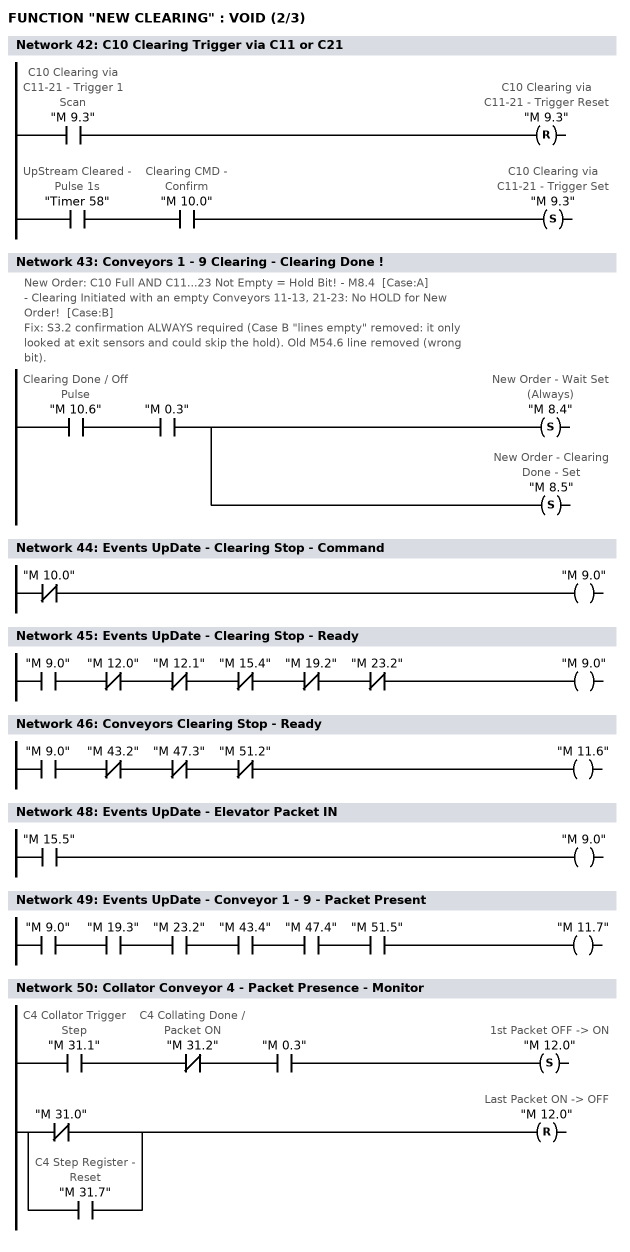

      A     "M 9.3"; // C10 Clearing via C11-21 - Trigger 1 Scan
      R     "M 9.3"; // C10 Clearing via C11-21 - Trigger Reset
//;
      A     "Timer 58"; // UpStream Cleared - Pulse 1s
      A     "M 10.0"; // Clearing CMD - Confirm
      S     "M 9.3"; // C10 Clearing via C11-21 - Trigger Set
NETWORK
TITLE =Conveyors 1 - 9 Clearing - Clearing Done !
//New Order: C10 Full AND C11...23 Not Empty = Hold Bit! - M8.4  [Case:A]
//
//- Clearing Initiated with an empty Conveyors 11-13, 21-23: No HOLD for New
//Order!  [Case:B]
//
//Fix: S3.2 confirmation ALWAYS required (Case B "lines empty" removed: it only
//looked at exit sensors and could skip the hold). Old M54.6 line removed (wrong
//bit).
      A     "M 10.6"; // Clearing Done / Off Pulse
      A     "M 0.3";
      S     "M 8.4"; // New Order - Wait Set (Always)
      S     "M 8.5"; // New Order - Clearing Done - Set
NETWORK
TITLE =Events UpDate - Clearing Stop - Command

      AN    "M 10.0";
      =     "M 9.0";
NETWORK
TITLE =Events UpDate - Clearing Stop - Ready

      A     "M 9.0";
      AN    "M 12.0";
      AN    "M 12.1";
      AN    "M 15.4";
      AN    "M 19.2";
      AN    "M 23.2";
      =     "M 9.0";
NETWORK
TITLE =Conveyors Clearing Stop - Ready

      A     "M 9.0";
      AN    "M 43.2";
      AN    "M 47.3";
      AN    "M 51.2";
      =     "M 11.6";
NETWORK
TITLE =New Order
//New Order : Start Filling Conveyors


NETWORK
TITLE =Events UpDate - Elevator Packet IN

      A     "M 15.5";
      =     "M 9.0";
NETWORK
TITLE =Events UpDate - Conveyor 1 - 9 - Packet Present

      A     "M 9.0";
      A     "M 19.3";
      A     "M 23.2";
      A     "M 43.4";
      A     "M 47.4";
      A     "M 51.5";
      =     "M 11.7";
NETWORK
TITLE =Collator Conveyor 4 - Packet Presence - Monitor

      A     "M 31.1"; // C4 Collator Trigger Step
      AN    "M 31.2"; // C4 Collating Done / Packet ON
      A     "M 0.3";
      S     "M 12.0"; // 1st Packet OFF -> ON
//;
      A(    ;
      ON    "M 31.0";
      O     "M 31.7"; // C4 Step Register - Reset
      )     ;
      R     "M 12.0"; // Last Packet ON -> OFF
NETWORK
TITLE =Collator Conveyor 10 - Packet Presence - Monitor
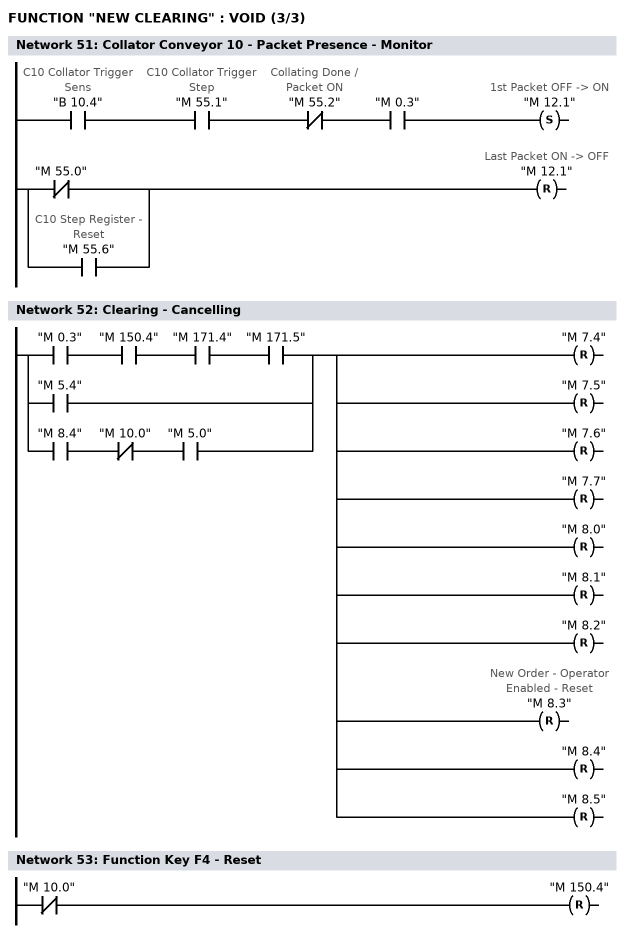

      A     "B 10.4"; // C10 Collator Trigger Sens
      A     "M 55.1"; // C10 Collator Trigger Step
      AN    "M 55.2"; // Collating Done / Packet ON
      A     "M 0.3";
      S     "M 12.1"; // 1st Packet OFF -> ON
//;
      A(    ;
      ON    "M 55.0";
      O     "M 55.6"; // C10 Step Register - Reset
      )     ;
      R     "M 12.1"; // Last Packet ON -> OFF
NETWORK
TITLE =Clearing - Cancelling

      A     "M 0.3";
      A     "M 150.4";
      A     "M 171.4";
      A     "M 171.5";
      O     "M 5.4";
      O(    ;
      A     "M 8.4";
      AN    "M 10.0";
      A     "M 5.0";
      )     ;
      R     "M 7.4";
      R     "M 7.5";
      R     "M 7.6";
      R     "M 7.7";
      R     "M 8.0";
      R     "M 8.1";
      R     "M 8.2";
      R     "M 8.3"; // New Order - Operator Enabled - Reset
      R     "M 8.4";
      R     "M 8.5";
NETWORK
TITLE =Function Key F4 - Reset

      AN    "M 10.0";
      R     "M 150.4";
END_FUNCTION

FUNCTION "NEW C0 + PUSHER 0" : VOID
TITLE =NEW FC912 (was FC1012) - Conveyor 0 & Pusher 0
NAME : 'Pos.1'
VERSION : 0.1


VAR_TEMP
  TIMER_RESET : BOOL ;
  MAIN_SERVICE_1_SW : BOOL ;
  CONV_0_SERVICE_FWD : BOOL ;
  CONV_0_SERVICE_REV : BOOL ;
  RESET_1 : BOOL ;
  RESET_2 : BOOL ;
  PUSHER_PUSH : BOOL ;
END_VAR
BEGIN
NETWORK
TITLE =Conveyor 0 - Service

      A     "HMI_DB".ALL_SERVICE_ENABLE_SW;
      A     "HMI_DB".CONVEYOR_0_SERVICE_SW;
      A     "HMI_DB".SERVICE_SW_1_STATUS;
      =     #MAIN_SERVICE_1_SW;
//;
      A     #MAIN_SERVICE_1_SW;
      O     "M 14.0";
      JNB   PUS0;
      A     "HMI_DB".HMI_ROLLER_TEST_FWD_SSW;
      FP    "FP 168.3";
      R     "HMI_DB".HMI_ROLLER_TEST_REV_SSW;
      =     #RESET_1;
//;
      A     "HMI_DB".HMI_ROLLER_TEST_REV_SSW;
      FP    "FP 168.4";
      R     "HMI_DB".HMI_ROLLER_TEST_FWD_SSW;
      =     #RESET_2;
//;
      A(    ;
      O     #RESET_1;
      O     #RESET_2;
      )     ;
      L     S5T#1S;
      SF    "Timer 110";
//;
      A     "HMI_DB".HMI_ROLLER_TEST_FWD_SSW;
      AN    "Timer 110";
      =     #CONV_0_SERVICE_FWD;
//;
      A     "HMI_DB".HMI_ROLLER_TEST_REV_SSW;
      AN    "Timer 110";
      =     #CONV_0_SERVICE_REV;
//;
      A     "HMI_DB".HMI_PUSHER_0_TEST_SSW;
      =     #PUSHER_PUSH;
//;
      AN    #MAIN_SERVICE_1_SW;
      R     "HMI_DB".HMI_ROLLER_TEST_FWD_SSW;
      R     "HMI_DB".HMI_ROLLER_TEST_REV_SSW;

PUS0: R     #CONV_0_SERVICE_FWD;
      R     #CONV_0_SERVICE_REV;
      R     #RESET_1;
      R     #RESET_2;
      R     #PUSHER_PUSH;
      FP    "FP 158.0";
      =     "M 14.0";
NETWORK
TITLE =Function Keys <F5 > on HMI - Reset
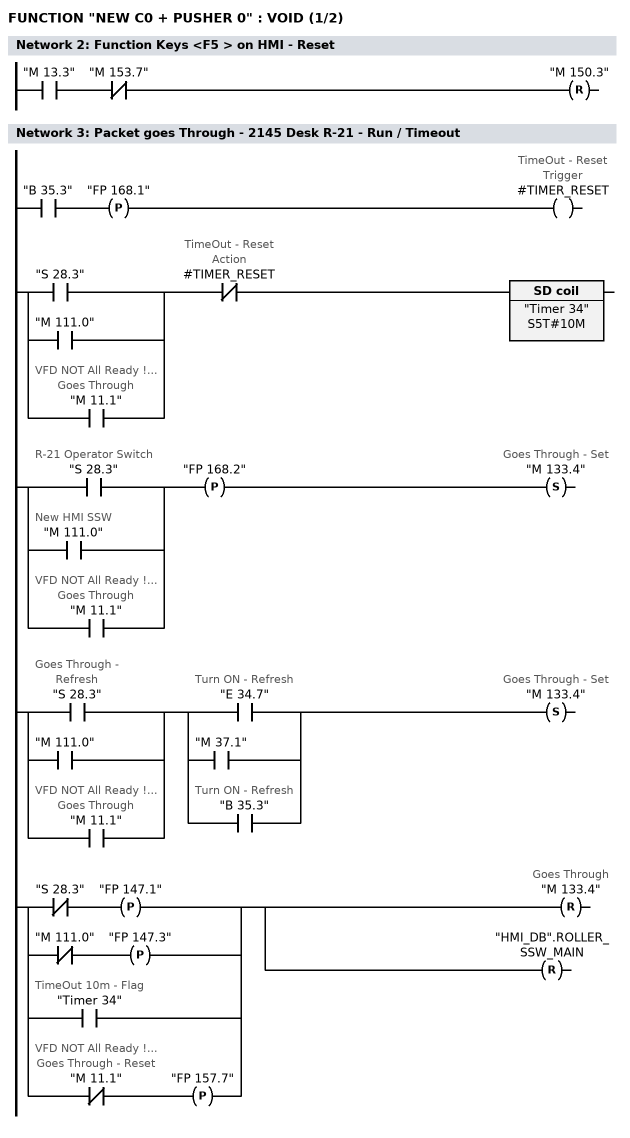

      A     "M 13.3";
      AN    "M 153.7";
      R     "M 150.3";
NETWORK
TITLE =Packet goes Through - 2145 Desk R-21 - Run / Timeout

      A     "B 35.3";
      FP    "FP 168.1";
      =     #TIMER_RESET; // TimeOut - Reset Trigger
//;
      A     "S 28.3";
      O     "M 111.0";
      O     "M 11.1"; // VFD NOT All Ready !... Goes Through
      AN    #TIMER_RESET; // TimeOut - Reset Action
      L     S5T#10M;
      SD    "Timer 34"; // TimeOut 10m
//;
      A     "S 28.3"; // R-21 Operator Switch
      O     "M 111.0"; // New HMI SSW
      O     "M 11.1"; // VFD NOT All Ready !... Goes Through
      FP    "FP 168.2"; // Turn ON - Pulse
      S     "M 133.4"; // Goes Through - Set
//;
      A     "S 28.3"; // Goes Through - Refresh
      O     "M 111.0";
      O     "M 11.1"; // VFD NOT All Ready !... Goes Through
      A(    ;
      O     "E 34.7"; // Turn ON - Refresh
      O     "M 37.1";
      O     "B 35.3"; // Turn ON - Refresh
      )     ;
      S     "M 133.4"; // Goes Through - Set
//;
      A(    ;
      O(    ;
      AN    "S 28.3";
      FP    "FP 147.1"; // Turn OFF - Pulse
      )     ;
      O(    ;
      AN    "M 111.0";
      FP    "FP 147.3"; // Turn OFF - Pulse
      O     "Timer 34"; // TimeOut 10m - Flag
      )     ;
      O(    ;
      AN    "M 11.1"; // VFD NOT All Ready !... Goes Through - Reset
      FP    "FP 157.7";
      )     ;
      )     ;
      R     "M 133.4"; // Goes Through
      R     "HMI_DB".ROLLER_SSW_MAIN;
NETWORK
TITLE =
//
//      A     "E 2.4"
//      S     "M 33.0"                    // Solid Detected ?
////;
//      A     "M 33.0"                    // Delay Timer - Start
//      L     S5T#300MS
//      SD    "Timer 26"                  // Debouncer 300mS
////;
//      A     "Timer 26"                  // Delayed Test Pulse
//      AN    "E 2.4"                     // Foul Detection
//      R     "M 33.0"                    // Not Detected !
////;
//      A     "Timer 26"                  // Delayed Test Pulse
//      A     "M 33.0"                    // Detection Comfirm !
//      =     "M 33.1"                    // Packet Height OK
//      R     "M 33.0"                    // Reset
//


NETWORK
TITLE =Packet Height - Sensing / Debouncing
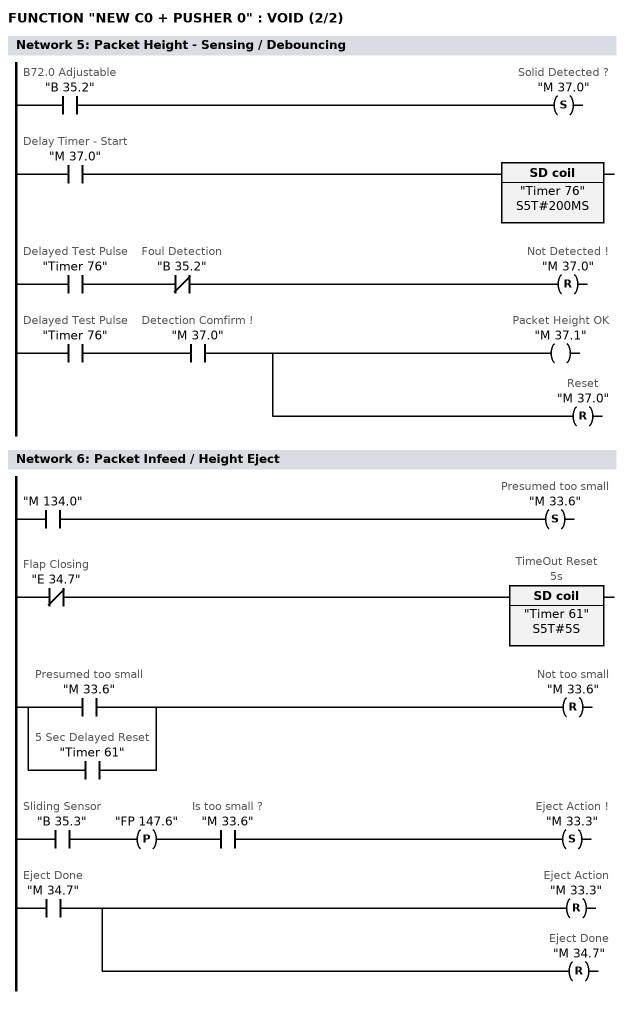

      A     "B 35.2"; // B72.0 Adjustable
      S     "M 37.0"; // Solid Detected ?
//;
      A     "M 37.0"; // Delay Timer - Start
      L     S5T#200MS;
      SD    "Timer 76"; // Debouncer 300mS
//;
      A     "Timer 76"; // Delayed Test Pulse
      AN    "B 35.2"; // Foul Detection
      R     "M 37.0"; // Not Detected !
//;
      A     "Timer 76"; // Delayed Test Pulse
      A     "M 37.0"; // Detection Comfirm !
      =     "M 37.1"; // Packet Height OK
      R     "M 37.0"; // Reset
NETWORK
TITLE =Packet Infeed / Height Eject

      A     "M 134.0";
      S     "M 33.6"; // Presumed too small
//;
      AN    "E 34.7"; // Flap Closing
      L     S5T#5S; // TimeOut Reset 5s
      SD    "Timer 61";
//;
      A     "M 33.6"; // Presumed too small
//    A     "M 33.1"                    // Packet Height OK ?
      O     "Timer 61"; // 5 Sec Delayed Reset
      R     "M 33.6"; // Not too small
//;
      A     "B 35.3"; // Sliding Sensor
      FP    "FP 147.6";
      A     "M 33.6"; // Is too small ?
      S     "M 33.3"; // Eject Action !
//;
      A     "M 34.7"; // Eject Done
      R     "M 33.3"; // Eject Action
      R     "M 34.7"; // Eject Done
NETWORK
TITLE =Eject Comfirmation

      A     "M 13.0";
      JNB   OUT1;

      A     "B 35.3";
      AN    "M 132.6"; // Not Triggered by Pusher
      S     "M 34.3"; // Eject Step 1
//;
      A     "B 35.4";
      AN    "M 132.6"; // Not Triggered by Pusher
      S     "M 34.4"; // Eject Step 2
//;
      A     "K 62.0"; // Conveyor 0 - Running
      A     "M 153.7";
      A     "M 34.3"; // Eject Step 1
      A     "M 34.4"; // Eject Step 2
      S     "M 34.5"; // Eject Step 3
//;
      A     "M 34.5"; // Eject Step 3
      AN    "B 35.4"; // Eject Step 4
      S     "M 34.7"; // Eject Done
      R     "M 34.3"; // Eject Step 1 - Reset
      R     "M 34.4"; // Eject Step 2 - Reset
      R     "M 34.5"; // Eject Step 3 - Reset
      R     "M 33.3"; // Eject Action - Reset
//;
      A     "M 132.5"; // Reset with Pusher Extend
      A     "B 35.4";
      R     "M 34.3"; // Eject Step 1 - Reset
      R     "M 34.4"; // Eject Step 2 - Reset
      R     "M 34.5"; // Eject Step 3 - Reset
      R     "M 33.3"; // Eject Action - Reset

OUT1: CLR   ;
NETWORK
TITLE =Packet goes Through - Conveyor 0 Man Run - LAUER F5
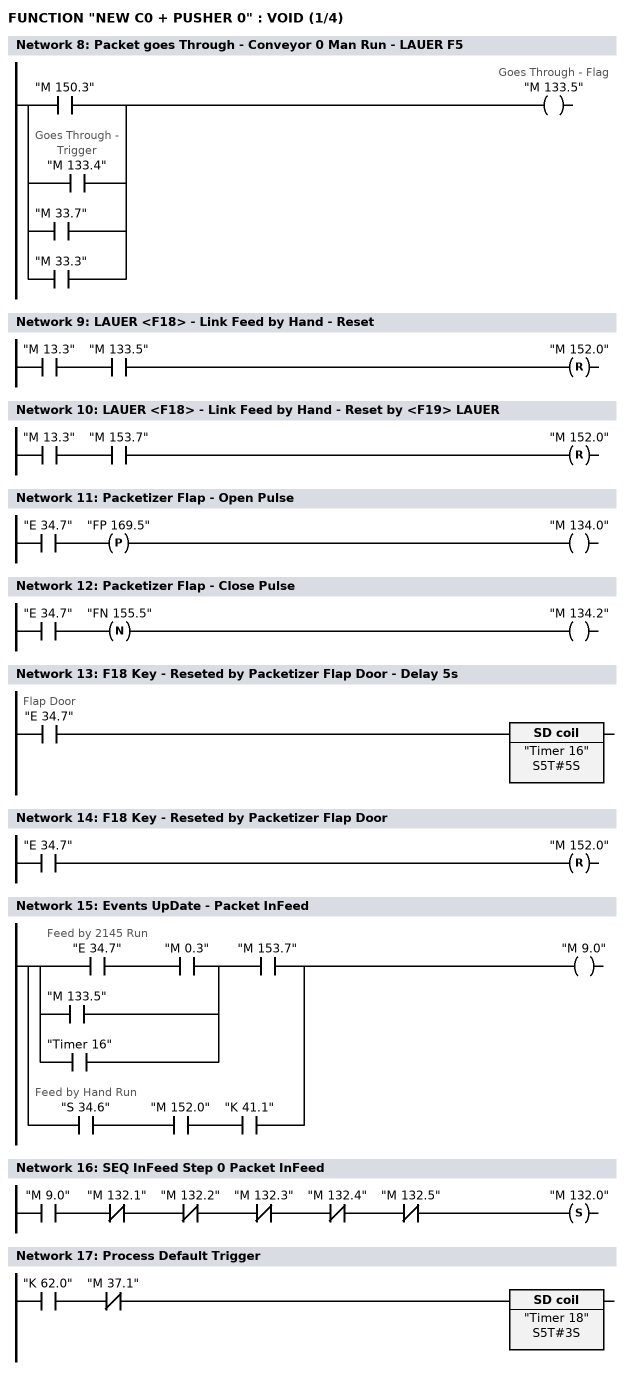

      O     "M 150.3";
      O     "M 133.4"; // Goes Through - Trigger
      O     "M 33.7";
      O     "M 33.3";
      =     "M 133.5"; // Goes Through - Flag
NETWORK
TITLE =LAUER <F18> - Link Feed by Hand - Reset

      A     "M 13.3";
      A     "M 133.5";
      R     "M 152.0";
NETWORK
TITLE =LAUER <F18> - Link Feed by Hand - Reset by <F19> LAUER

      A     "M 13.3";
      A     "M 153.7";
      R     "M 152.0";
NETWORK
TITLE =Packetizer Flap - Open Pulse

      A     "E 34.7";
      FP    "FP 169.5";
      =     "M 134.0";
NETWORK
TITLE =Packetizer Flap - Close Pulse

      A     "E 34.7";
      FN    "FN 155.5";
      =     "M 134.2";
NETWORK
TITLE =F18 Key - Reseted by Packetizer Flap Door - Delay 5s

      A     "E 34.7"; // Flap Door
      L     S5T#5S;
      SD    "Timer 16"; // Setup Mode Trigger
NETWORK
TITLE =F18 Key - Reseted by Packetizer Flap Door

      A     "E 34.7";
      R     "M 152.0";
NETWORK
TITLE =Events UpDate - Packet InFeed

      A(    ;
      A     "E 34.7"; // Feed by 2145 Run
      A     "M 0.3";
      O     "M 133.5";
      O     "Timer 16";
      A     "M 153.7";
      O     ;
      A     "S 34.6"; // Feed by Hand Run
      A     "M 152.0";
      A     "K 41.1";
      )     ;
      =     "M 9.0";
NETWORK
TITLE =SEQ InFeed Step 0 Packet InFeed

      A     "M 9.0";
      AN    "M 132.1";
      AN    "M 132.2";
      AN    "M 132.3";
      AN    "M 132.4";
      AN    "M 132.5";
      S     "M 132.0";
NETWORK
TITLE =Process Default Trigger

      A     "K 62.0";
      AN    "M 37.1";
      L     S5T#3S;
      SD    "Timer 18";
NETWORK
TITLE =Events UpDate
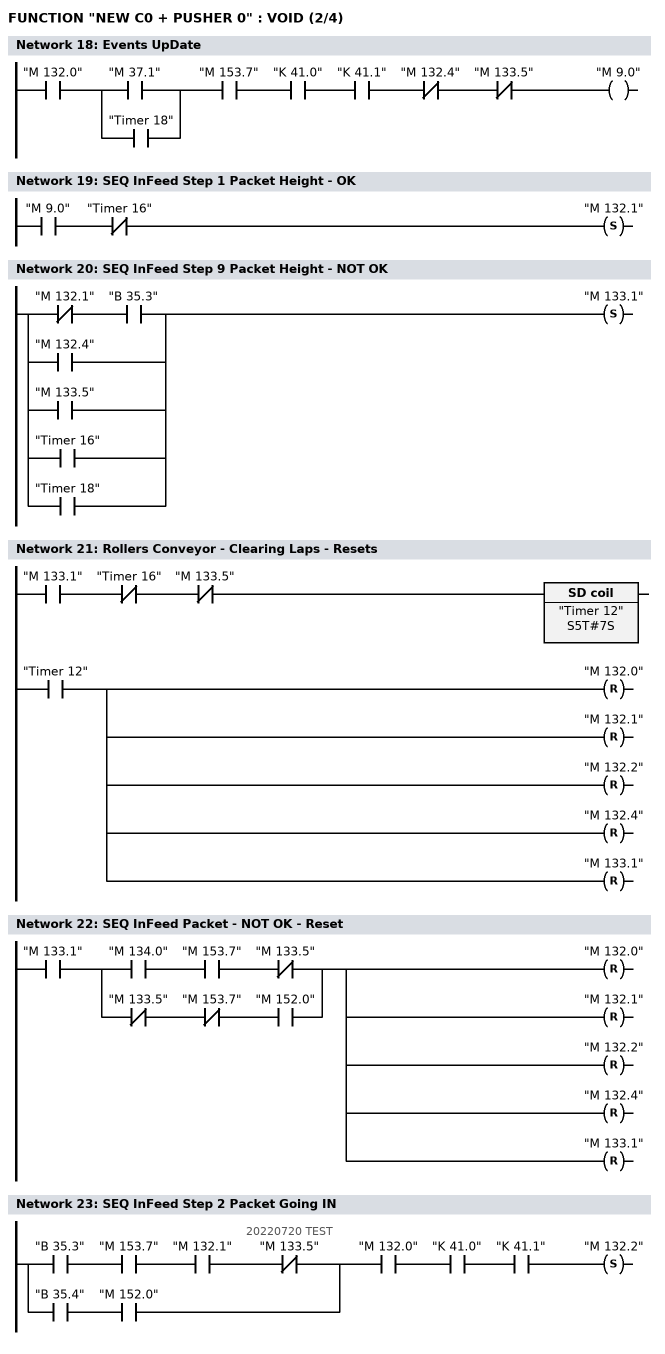

      A     "M 132.0";
      A(    ;
      O     "M 37.1";
      O     "Timer 18";
      )     ;
      A     "M 153.7";
      A     "K 41.0";
      A     "K 41.1";
      AN    "M 132.4";
      AN    "M 133.5";
      =     "M 9.0";
NETWORK
TITLE =SEQ InFeed Step 1 Packet Height - OK

      A     "M 9.0";
      AN    "Timer 16";
      S     "M 132.1";
NETWORK
TITLE =SEQ InFeed Step 9 Packet Height - NOT OK

      AN    "M 132.1";
      A     "B 35.3";
      O     "M 132.4";
      O     "M 133.5";
      O     "Timer 16";
      O     "Timer 18";
      S     "M 133.1";
NETWORK
TITLE =Rollers Conveyor - Clearing Laps - Resets

      A     "M 133.1";
      AN    "Timer 16";
      AN    "M 133.5";
      L     S5T#7S;
      SD    "Timer 12";
//;
      A     "Timer 12";
      R     "M 132.0";
      R     "M 132.1";
      R     "M 132.2";
      R     "M 132.4";
      R     "M 133.1";
NETWORK
TITLE =SEQ InFeed Packet - NOT OK - Reset

      A     "M 133.1";
      A(    ;
      A     "M 134.0";
      A     "M 153.7";
      AN    "M 133.5";
      O     ;
      AN    "M 133.5";
      AN    "M 153.7";
      A     "M 152.0";
      )     ;
      R     "M 132.0";
      R     "M 132.1";
      R     "M 132.2";
      R     "M 132.4";
      R     "M 133.1";
NETWORK
TITLE =SEQ InFeed Step 2 Packet Going IN

      A(    ;
      A     "B 35.3";
      A     "M 153.7";
      A     "M 132.1";
      AN    "M 133.5"; // 20220720 TEST
      O     ;
      A     "B 35.4";
      A     "M 152.0";
      )     ;
      A     "M 132.0";
      A     "K 41.0";
      A     "K 41.1";
      S     "M 132.2";
NETWORK
TITLE =SEQ InFeed Step 3 Conveyor Stop
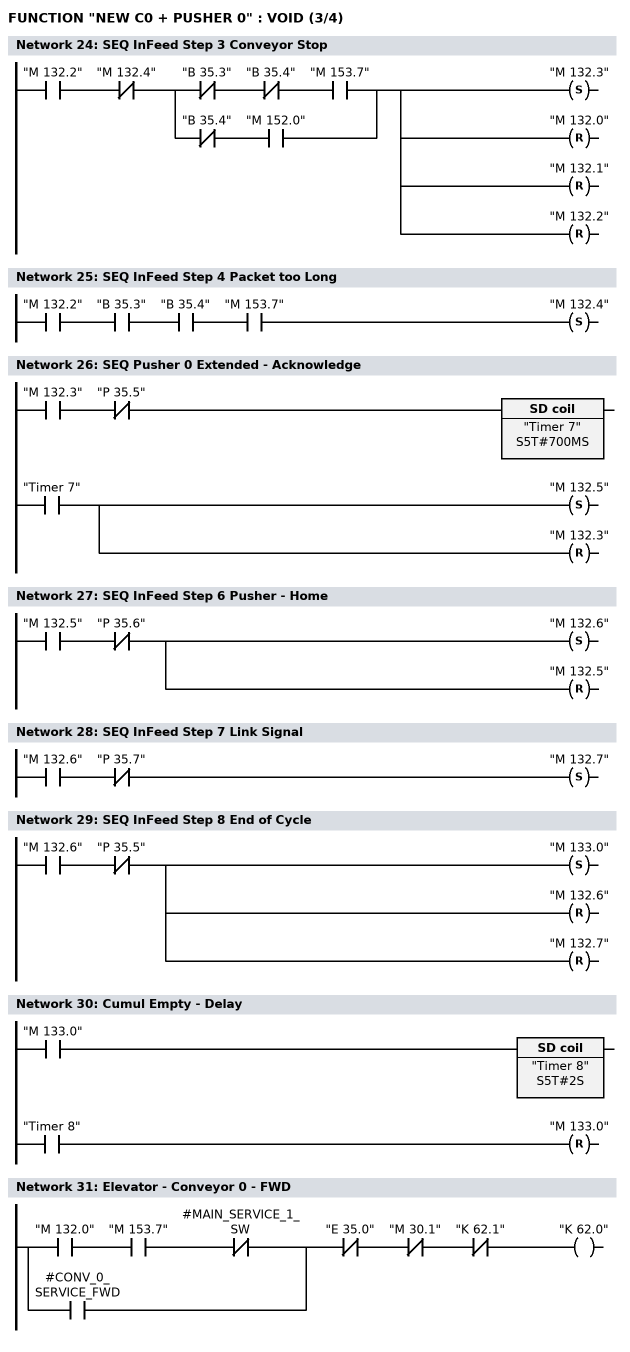

      A     "M 132.2";
      AN    "M 132.4";
      A(    ;
      AN    "B 35.3";
      AN    "B 35.4";
      A     "M 153.7";
      O     ;
      AN    "B 35.4";
      A     "M 152.0";
      )     ;
      S     "M 132.3";
      R     "M 132.0";
      R     "M 132.1";
      R     "M 132.2";
NETWORK
TITLE =SEQ InFeed Step 4 Packet too Long

      A     "M 132.2";
      A     "B 35.3";
      A     "B 35.4";
      A     "M 153.7";
      S     "M 132.4";
NETWORK
TITLE =SEQ Pusher 0 Extended - Acknowledge

      A     "M 132.3";
      AN    "P 35.5";
      L     S5T#700MS;
      SD    "Timer 7";
//;
      A     "Timer 7";
      S     "M 132.5";
      R     "M 132.3";
NETWORK
TITLE =SEQ InFeed Step 6 Pusher - Home

      A     "M 132.5";
      AN    "P 35.6";
      S     "M 132.6";
      R     "M 132.5";
NETWORK
TITLE =SEQ InFeed Step 7 Link Signal

      A     "M 132.6";
      AN    "P 35.7";
      S     "M 132.7";
NETWORK
TITLE =SEQ InFeed Step 8 End of Cycle

      A     "M 132.6";
      AN    "P 35.5";
      S     "M 133.0";
      R     "M 132.6";
      R     "M 132.7";
NETWORK
TITLE =Cumul Empty - Delay

      A     "M 133.0";
      L     S5T#2S;
      SD    "Timer 8";
//;
      A     "Timer 8";
      R     "M 133.0";
NETWORK
TITLE =Elevator - Conveyor 0 - FWD

      A(    ;
      A     "M 132.0";
      A     "M 153.7";
      AN    #MAIN_SERVICE_1_SW;
      O     #CONV_0_SERVICE_FWD;
      )     ;
      AN    "E 35.0";
      AN    "M 30.1";
      AN    "K 62.1";
      =     "K 62.0";
NETWORK
TITLE =Elevator - Conveyor 0 - REV
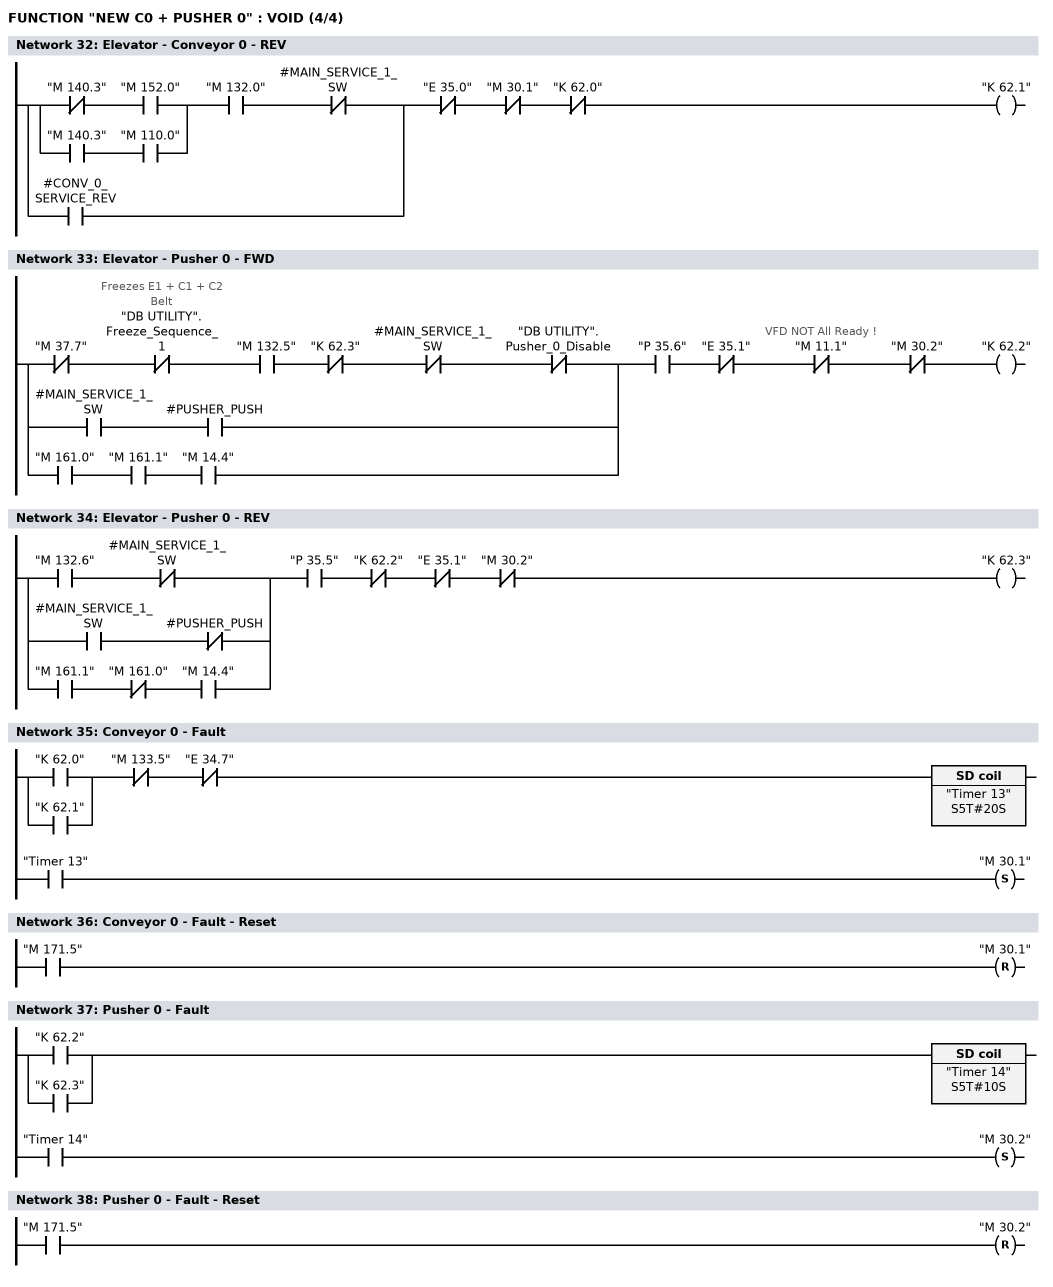

      A(    ;
      A(    ;
      AN    "M 140.3";
      A     "M 152.0";
      O     ;
      A     "M 140.3";
      A     "M 110.0";
      )     ;
      A     "M 132.0";
//     A     "M 152.0"
      AN    #MAIN_SERVICE_1_SW;
      O     #CONV_0_SERVICE_REV;
      )     ;
      AN    "E 35.0";
      AN    "M 30.1";
      AN    "K 62.0";
      =     "K 62.1";
NETWORK
TITLE =Elevator - Pusher 0 - FWD

      A(    ;
      AN    "M 37.7";
      AN    "DB UTILITY".Freeze_Sequence_1; //  Freezes E1 + C1 + C2 Belt
      A     "M 132.5";
      AN    "K 62.3";
      AN    #MAIN_SERVICE_1_SW;
      AN    "DB UTILITY".Pusher_0_Disable;
      O(    ;
      A     #MAIN_SERVICE_1_SW;
      A     #PUSHER_PUSH;
      )     ;
      O     ;
      A     "M 161.0";
      A     "M 161.1";
      A     "M 14.4";
      )     ;
      A     "P 35.6";
      AN    "E 35.1";
      AN    "M 11.1"; // VFD NOT All Ready !
      AN    "M 30.2";
      =     "K 62.2";
NETWORK
TITLE =Elevator - Pusher 0 - REV

      A(    ;
      A     "M 132.6";
      AN    #MAIN_SERVICE_1_SW;
      O(    ;
      A     #MAIN_SERVICE_1_SW;
      AN    #PUSHER_PUSH;
      )     ;
      O     ;
      A     "M 161.1";
      AN    "M 161.0";
      A     "M 14.4";
      )     ;
      A     "P 35.5";
      AN    "K 62.2";
      AN    "E 35.1";
      AN    "M 30.2";
      =     "K 62.3";
NETWORK
TITLE =Conveyor 0 - Fault

      A(    ;
      O     "K 62.0";
      O     "K 62.1";
      )     ;
      AN    "M 133.5";
      AN    "E 34.7";
      L     S5T#20S;
      SD    "Timer 13";
//;
      A     "Timer 13";
      S     "M 30.1";
NETWORK
TITLE =Conveyor 0 - Fault - Reset

      A     "M 171.5";
      R     "M 30.1";
NETWORK
TITLE =Pusher 0 - Fault

      A(    ;
      O     "K 62.2";
      O     "K 62.3";
      )     ;
      L     S5T#10S;
      SD    "Timer 14";
//;
      A     "Timer 14";
      S     "M 30.2";
NETWORK
TITLE =Pusher 0 - Fault - Reset

      A     "M 171.5";
      R     "M 30.2";
END_FUNCTION

FUNCTION "NEW ELEVATOR + PUSHER 1" : VOID
TITLE =NEW FC916 (was FC1016) - Elevator + Pusher 1 Pos.2
//
NAME : POS_2
VERSION : 0.0


VAR_TEMP
  ELEVATOR_UP_OUT : BOOL ;
  ELEVATOR_DN_OUT : BOOL ;
  MAIN_SERVICE_1_SW : BOOL ;
  ELEVATOR_SERVICE_SW : BOOL ;
  ELEVATOR_DN_PB : BOOL ;
  ELEVATOR_UP_PB : BOOL ;
  ELEVATOR_ROUNDTRIP : BOOL ;
  PUSHER_PUSH : BOOL ;
  INITIALISATION : BOOL ;
  BRAKE_RELEASE_OK : BOOL ;
  BRAKE_CONTACTOR_KO : BOOL ;
END_VAR
BEGIN
NETWORK
TITLE =Elevator - Health OK
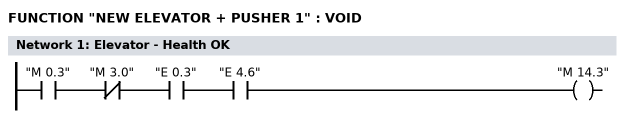

      A     "M 0.3";
      AN    "M 3.0";
      A     "E 0.3";
      A     "E 4.6";
      =     "M 14.3";
NETWORK
TITLE =Elevator - Service

      A     "HMI_DB".ALL_SERVICE_ENABLE_SW;
      A     "HMI_DB".ELEVATOR_SERVICE_SW;
      A     "HMI_DB".SERVICE_SW_1_STATUS;
      =     #MAIN_SERVICE_1_SW;
//;
      A     #MAIN_SERVICE_1_SW;
      O     "M 14.1";
      JNB   PUS1;
      A     "HMI_DB".HMI_ELEVATOR_SERVICE_SSW;
      =     #ELEVATOR_SERVICE_SW;
      S     "DB UTILITY".Pusher_0_Disable;
//;
      A     #ELEVATOR_SERVICE_SW;
      A(    ;
      A     "HMI_DB".HMI_ELEVATOR_TEST_DN_SSW;
      )     ;
      =     #ELEVATOR_DN_PB;
//;
      A     #ELEVATOR_SERVICE_SW;
      A(    ;
      A     "HMI_DB".HMI_ELEVATOR_TEST_UP_SSW;
      )     ;
      =     #ELEVATOR_UP_PB;
//;
      A     #MAIN_SERVICE_1_SW;
      AN    #ELEVATOR_SERVICE_SW;
      A     "HMI_DB".ELEVATOR_ROUND_TRIP_SSW;
      =     #ELEVATOR_ROUNDTRIP;
//;
      A     "HMI_DB".HMI_PUSHER_1_TEST_SSW;
      =     #PUSHER_PUSH;
//;
      AN    #MAIN_SERVICE_1_SW;
      R     "HMI_DB".HMI_ELEVATOR_SERVICE_SSW;
      R     "HMI_DB".HMI_ELEVATOR_TEST_DN_SSW;
      R     "HMI_DB".HMI_ELEVATOR_TEST_UP_SSW;
      R     "DB UTILITY".Pusher_0_Disable;

PUS1: R     #ELEVATOR_SERVICE_SW;
      R     #ELEVATOR_DN_PB;
      R     #ELEVATOR_UP_PB;
      R     #ELEVATOR_ROUNDTRIP;
      R     #PUSHER_PUSH;
      FP    "FP 158.1";
      =     "M 14.1";
//;
      A     "HMI_DB".SERVICE_INIT_PB;
      A     #ELEVATOR_SERVICE_SW;
      A     #MAIN_SERVICE_1_SW;
      =     #INITIALISATION;
NETWORK
TITLE =Elevator - Manual Run - Conditions
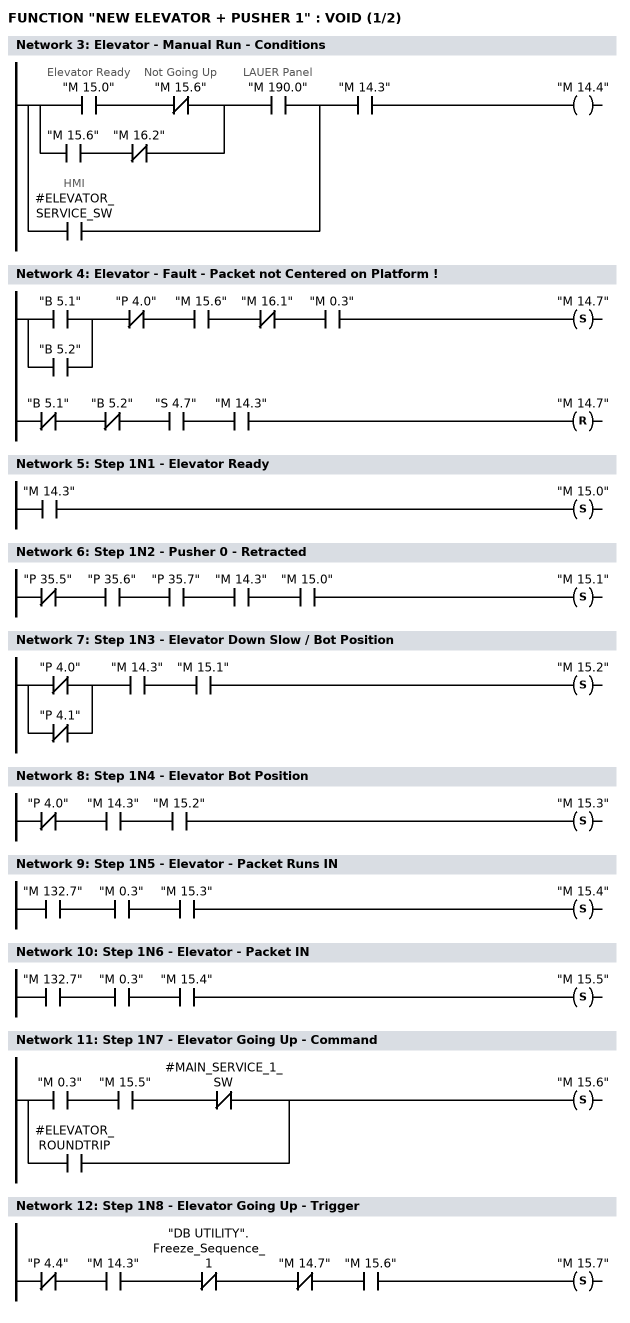

      A(    ;
      A     "M 15.0"; // Elevator Ready
      AN    "M 15.6"; // Not Going Up
      O     ; // or
      A     "M 15.6";
      AN    "M 16.2";
      )     ;
      A     "M 190.0"; // LAUER Panel
      O     #ELEVATOR_SERVICE_SW; // HMI
      A     "M 14.3";
      =     "M 14.4";
NETWORK
TITLE =Elevator - Fault - Packet not Centered on Platform !

      A(    ;
      O     "B 5.1";
      O     "B 5.2";
      )     ;
      AN    "P 4.0";
      A     "M 15.6";
      AN    "M 16.1";
      A     "M 0.3";
      S     "M 14.7";
//;
      AN    "B 5.1";
      AN    "B 5.2";
      A     "S 4.7";
      A     "M 14.3";
      R     "M 14.7";
NETWORK
TITLE =Step 1N1 - Elevator Ready

      A     "M 14.3";
      S     "M 15.0";
NETWORK
TITLE =Step 1N2 - Pusher 0 - Retracted

      AN    "P 35.5";
      A     "P 35.6";
      A     "P 35.7";
      A     "M 14.3";
      A     "M 15.0";
      S     "M 15.1";
NETWORK
TITLE =Step 1N3 - Elevator Down Slow / Bot Position

      A(    ;
      ON    "P 4.0";
      ON    "P 4.1";
      )     ;
      A     "M 14.3";
      A     "M 15.1";
      S     "M 15.2";
NETWORK
TITLE =Step 1N4 - Elevator Bot Position

      AN    "P 4.0";
      A     "M 14.3";
      A     "M 15.2";
      S     "M 15.3";
NETWORK
TITLE =Step 1N5 - Elevator - Packet Runs IN

      A     "M 132.7";
      A     "M 0.3";
      A     "M 15.3";
      S     "M 15.4";
NETWORK
TITLE =Step 1N6 - Elevator - Packet IN

      A     "M 132.7";
      A     "M 0.3";
      A     "M 15.4";
      S     "M 15.5";
NETWORK
TITLE =Step 1N7 - Elevator Going Up - Command

      A     "M 0.3";
      A     "M 15.5";
      AN    #MAIN_SERVICE_1_SW;
      O     #ELEVATOR_ROUNDTRIP;
      S     "M 15.6";
NETWORK
TITLE =Step 1N8 - Elevator Going Up - Trigger

      AN    "P 4.4";
      A     "M 14.3";
      AN    "DB UTILITY".Freeze_Sequence_1;
      AN    "M 14.7";
      A     "M 15.6";
      S     "M 15.7";
NETWORK
TITLE =Step 1N9 - Elevator Going Up - Slow
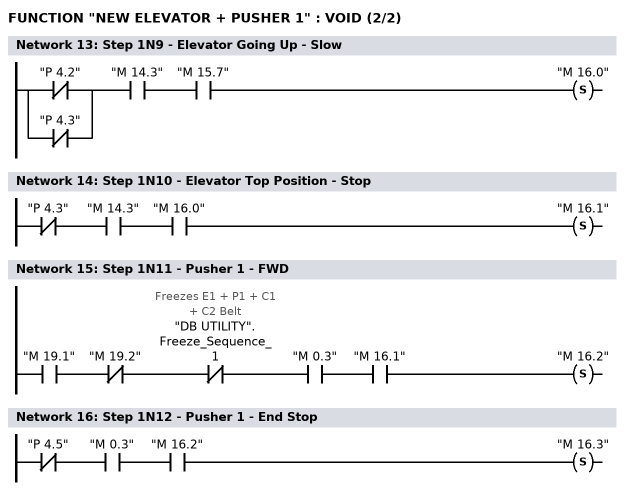

      A(    ;
      ON    "P 4.2";
      ON    "P 4.3";
      )     ;
      A     "M 14.3";
      A     "M 15.7";
      S     "M 16.0";
NETWORK
TITLE =Step 1N10 - Elevator Top Position - Stop

      AN    "P 4.3";
      A     "M 14.3";
      A     "M 16.0";
      S     "M 16.1";
NETWORK
TITLE =Step 1N11 - Pusher 1 - FWD

      A     "M 19.1";
      AN    "M 19.2";
      AN    "DB UTILITY".Freeze_Sequence_1; //  Freezes E1 + P1 + C1 + C2 Belt
      A     "M 0.3";
      A     "M 16.1";
      S     "M 16.2";
NETWORK
TITLE =Step 1N12 - Pusher 1 - End Stop

      AN    "P 4.5";
      A     "M 0.3";
      A     "M 16.2";
      S     "M 16.3";
NETWORK
TITLE =Soft Timer 15 Reset

      A     "M 16.3";
      AN    "M 16.4";
      A     "M 14.3";
      A     "M 0.3";
      JCN   R151;
      JU    E151;

R151: L     L#0;
      T     "DB UTILITY".T15_ET;
      R     "DB UTILITY".T15_DN;

E151: NOP   0;

NETWORK
TITLE =Soft Timer 15 Add

      A     "M 16.3";
      AN    "M 16.4";
      A     "M 14.3";
      A     "M 0.3";
      AN    "DB UTILITY".Freeze_Sequence_1;
      AN    "DB UTILITY".T15_DN;
      JCN   E152;

      L     "DB UTILITY".T15_ET;
      L     "DB UTILITY".Scan_Cycle_Previous;
      ITD   ;
      +D    ;
      T     "DB UTILITY".T15_ET;

E152: NOP   0;

NETWORK
TITLE =Soft Timer 15 Done 100mS
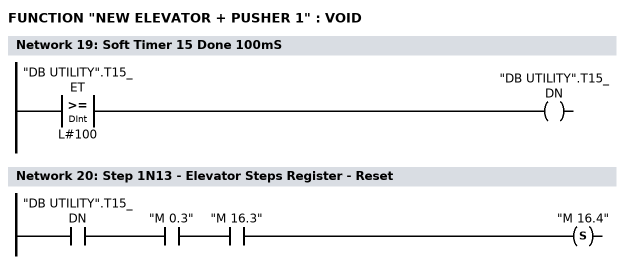

      L     "DB UTILITY".T15_ET;
      L     L#100;
      >=D   ;
      =     "DB UTILITY".T15_DN;

NETWORK
TITLE =Step 1N13 - Elevator Steps Register - Reset

      A     "DB UTILITY".T15_DN;
      A     "M 0.3";
      A     "M 16.3";
      S     "M 16.4";
NETWORK
TITLE =Elevator Steps Register - Reset

      A(    ;
      A     "M 190.0";
      A     "M 171.4";
      A     "M 171.5";
      O     "M 16.4";
      O     #INITIALISATION;
      O     "DB UTILITY".Elevator_Disable;
      )     ;
      A     "M 0.3";
      JC    M001;
      JU    M002;

M001: L     W#16#0;
      T     "MW 15";

M002: CLR   ;
NETWORK
TITLE =Trans System - Ready -> Tuber 2145
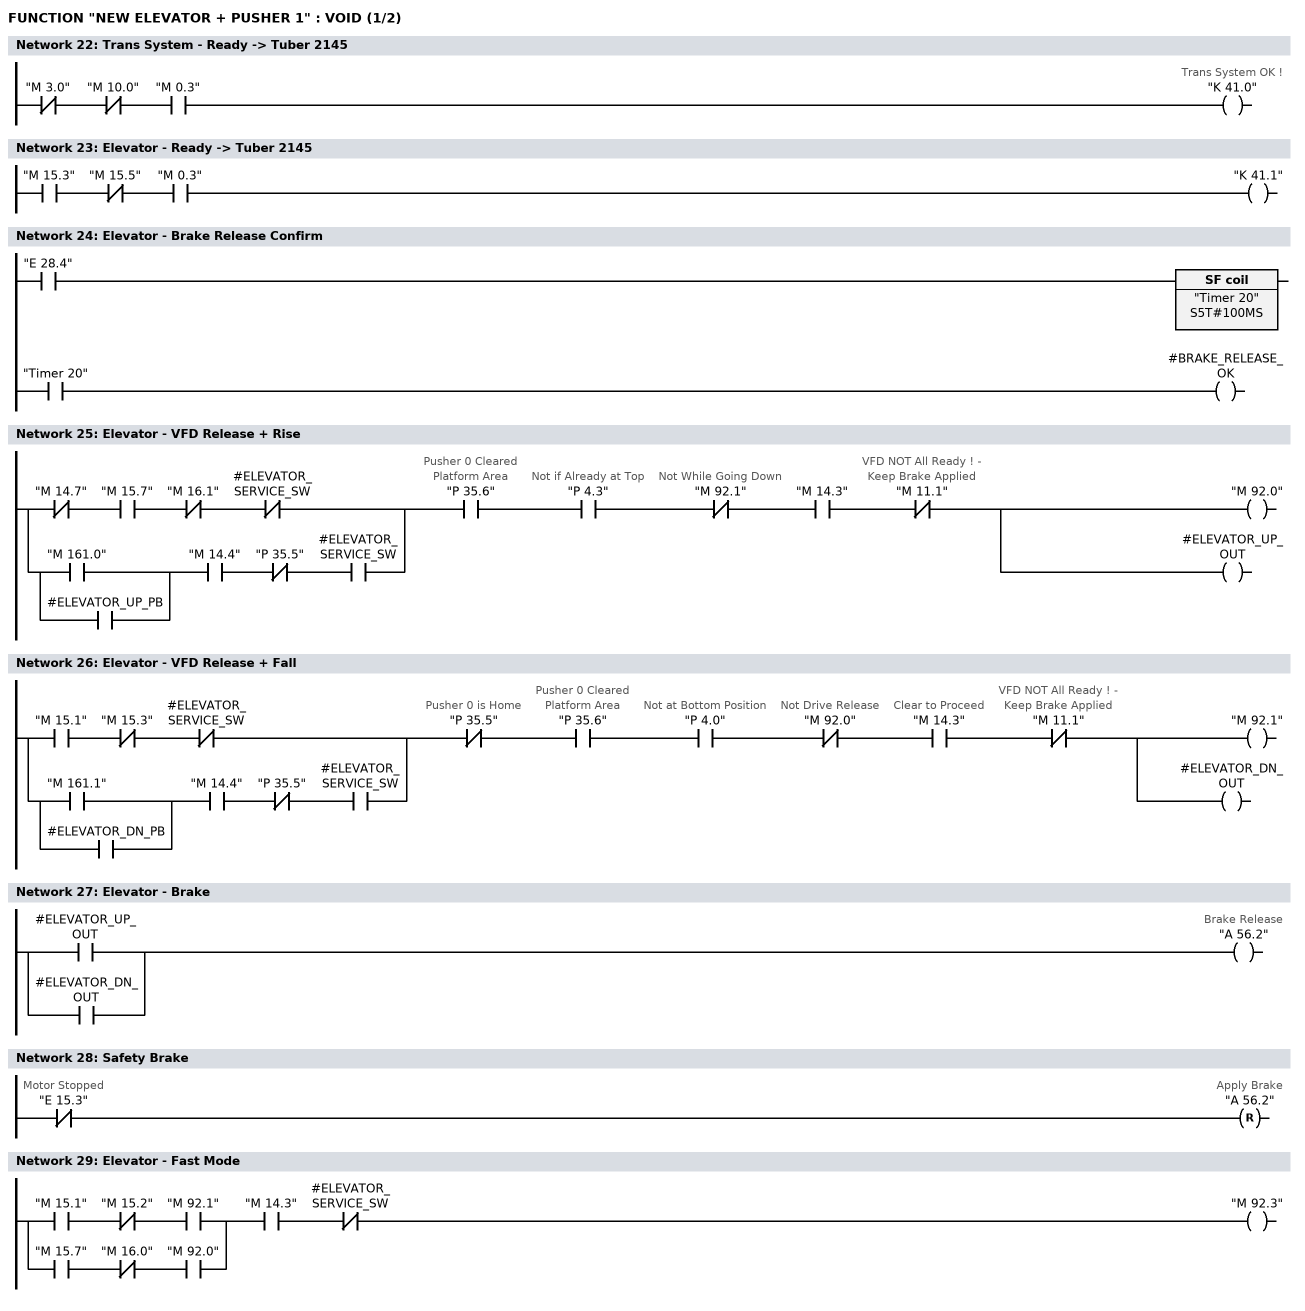

      AN    "M 3.0";
      AN    "M 10.0";
      A     "M 0.3";
      =     "K 41.0"; // Trans System OK !
NETWORK
TITLE =Elevator - Ready -> Tuber 2145

      A     "M 15.3";
      AN    "M 15.5";
      A     "M 0.3";
      =     "K 41.1";
NETWORK
TITLE =Elevator - Brake Release Confirm

      A     "E 28.4";
      L     S5T#100MS;
      SF    "Timer 20";
//;
      A     "Timer 20";
      =     #BRAKE_RELEASE_OK;
NETWORK
TITLE =Elevator - VFD Release + Rise

      A(    ;
      AN    "M 14.7";
      A     "M 15.7";
      AN    "M 16.1";
      AN    #ELEVATOR_SERVICE_SW;
      O     ;
      A(    ;
      O     "M 161.0";
      O     #ELEVATOR_UP_PB;
      )     ;
      A     "M 14.4";
      AN    "P 35.5";
      A     #ELEVATOR_SERVICE_SW;
      )     ;
      A     "P 35.6"; // Pusher 0 Cleared Platform Area
      A     "P 4.3"; // Not if Already at Top
      AN    "M 92.1"; // Not While Going Down
      A     "M 14.3";
      AN    "M 11.1"; // VFD NOT All Ready ! - Keep Brake Applied
      =     "M 92.0";
      =     #ELEVATOR_UP_OUT;
NETWORK
TITLE =Elevator - VFD Release + Fall

      A(    ;
      A     "M 15.1";
      AN    "M 15.3";
      AN    #ELEVATOR_SERVICE_SW;
      O     ;
      A(    ;
      O     "M 161.1";
      O     #ELEVATOR_DN_PB;
      )     ;
      A     "M 14.4";
      AN    "P 35.5";
      A     #ELEVATOR_SERVICE_SW;
      )     ;
      AN    "P 35.5"; // Pusher 0 is Home
      A     "P 35.6"; // Pusher 0 Cleared Platform Area
      A     "P 4.0"; // Not at Bottom Position
      AN    "M 92.0"; // Not Drive Release
      A     "M 14.3"; // Clear to Proceed
      AN    "M 11.1"; // VFD NOT All Ready ! - Keep Brake Applied
      =     "M 92.1";
      =     #ELEVATOR_DN_OUT;
NETWORK
TITLE =Elevator - Brake

      A(    ;
      O     #ELEVATOR_UP_OUT;
      O     #ELEVATOR_DN_OUT;
      )     ;
      =     "A 56.2"; // Brake Release
NETWORK
TITLE =Safety Brake

      AN    "E 15.3"; // Motor Stopped
      R     "A 56.2"; // Apply Brake
NETWORK
TITLE =Elevator - Fast Mode

      A(    ;
      A     "M 15.1";
      AN    "M 15.2";
      A     "M 92.1";
      O     ;
      A     "M 15.7";
      AN    "M 16.0";
      A     "M 92.0";
      )     ;
      A     "M 14.3";
      AN    #ELEVATOR_SERVICE_SW;
      =     "M 92.3";
NETWORK
TITLE =Elevator - Slow
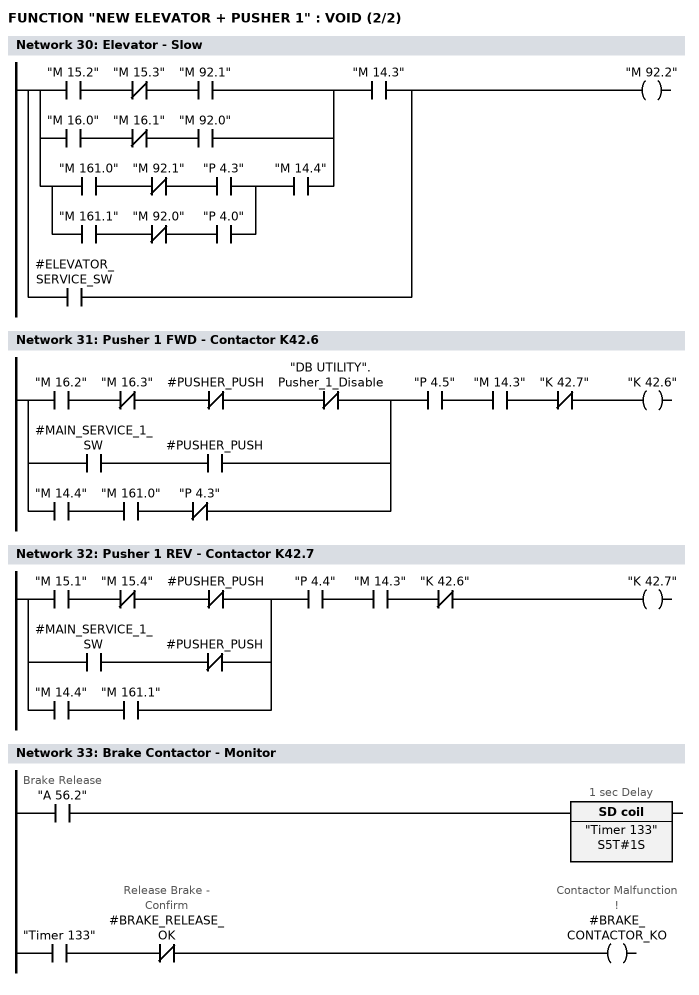

      A(    ;
      A     "M 15.2";
      AN    "M 15.3";
      A     "M 92.1";
      O     ;
      A     "M 16.0";
      AN    "M 16.1";
      A     "M 92.0";
      O     ;
      A(    ;
      A     "M 161.0";
      AN    "M 92.1";
      A     "P 4.3";
      O     ;
      A     "M 161.1";
      AN    "M 92.0";
      A     "P 4.0";
      )     ;
      A     "M 14.4";
      )     ;
      A     "M 14.3";
      O     #ELEVATOR_SERVICE_SW;
      =     "M 92.2";
NETWORK
TITLE =Pusher 1 FWD - Contactor K42.6

      A(    ;
      A     "M 16.2";
      AN    "M 16.3";
      AN    #PUSHER_PUSH;
      AN    "DB UTILITY".Pusher_1_Disable;
      O(    ;
      A     #MAIN_SERVICE_1_SW;
      A     #PUSHER_PUSH;
      )     ;
      O     ;
      A     "M 14.4";
      A     "M 161.0";
      AN    "P 4.3";
      )     ;
      A     "P 4.5";
      A     "M 14.3";
      AN    "K 42.7";
      =     "K 42.6";
NETWORK
TITLE =Pusher 1 REV - Contactor K42.7

      A(    ;
      A     "M 15.1";
      AN    "M 15.4";
      AN    #PUSHER_PUSH;
      O(    ;
      A     #MAIN_SERVICE_1_SW;
      AN    #PUSHER_PUSH;
      )     ;
      O     ;
      A     "M 14.4";
      A     "M 161.1";
      )     ;
      A     "P 4.4";
      A     "M 14.3";
      AN    "K 42.6";
      =     "K 42.7";
NETWORK
TITLE =Brake Contactor - Monitor

      A     "A 56.2"; // Brake Release
      L     S5T#1S; // 1 sec Delay
      SD    "Timer 133";
//;
      A     "Timer 133";
      AN    #BRAKE_RELEASE_OK; // Release Brake - Confirm
      =     #BRAKE_CONTACTOR_KO; // Contactor Malfunction !
NETWORK
TITLE =New Elevator VFD PARKER - Ready

      AN    "E 14.4"; // DRIVE TEST
      O     #BRAKE_CONTACTOR_KO; // Contactor Monitor = Contactor Malfunction !
      JCN   NFLT; // No fault
      S     "M 92.5"; // Set Fault Bit
      JU    OFF; // Turn Off
NETWORK
TITLE =New Elevator VFD with Dynamic Resistor - Go Up

NFLT: A     #ELEVATOR_UP_OUT; // VFD Release Command UP
      A     "M 92.3"; // Fast Speed Command
      AN    "M 92.5"; // Fault Bit
      AN    "M 11.1"; // VFD NOT All Ready !
      JCN   UPLO;
      S     "A 63.0"; // Release Drive - Go Up
      S     "A 63.2"; // Speed 2 / Speed 0.0
//;
      A     #BRAKE_RELEASE_OK; // Release Brake - Confirm
      JCN   END;
      =     "A 63.1"; // Speed 1
      =     "A 63.2"; // Speed 2 + Speed 1 = Fast
      R     "A 63.3"; // L = Forward (Up)
      JU    END;

UPLO: A     #ELEVATOR_UP_OUT; // VFD Release Command UP
      A     "M 92.2"; // Slow Speed Command
      AN    "M 92.5"; // Fault Bit
      AN    "M 11.1"; // VFD NOT All Ready !
      JCN   DNHI;
      S     "A 63.0"; // Release Drive - Go Up
      S     "A 63.2"; // Speed 2 / Speed 0.0
//;
      A     #BRAKE_RELEASE_OK; // Release Brake - Confirm
      JCN   END;
      =     "A 63.1"; // Speed 1
      R     "A 63.2"; // Speed 2 = Off
      R     "A 63.3"; // L = Forward (Up)
      JU    END;
NETWORK
TITLE =New Elevator VFD with Dynamic Resistor - Go Down

DNHI: A     #ELEVATOR_DN_OUT; // VFD Release Command DN
      A     "M 92.3"; // Fast Speed Command
      AN    "M 92.5"; // Fault Bit
      JCN   DNLO;
      S     "A 63.0"; // Release Drive - Go Dn
      S     "A 63.2"; // Speed 2 / Speed 0.0
//;
      A     #BRAKE_RELEASE_OK; // Release Brake - Confirm
      JCN   END;
      =     "A 63.1"; // Speed 1
      =     "A 63.2"; // Speed 2 + Speed 1 = Fast
      =     "A 63.3"; // H = Reverse (Dn)
      JU    END;

DNLO: A     #ELEVATOR_DN_OUT; // VFD Release Command DN
      A     "M 92.2"; // Slow Speed Command
      AN    "M 92.5"; // Fault Bit
      JCN   OFF;
      S     "A 63.0"; // Release Drive - Go Dn
      S     "A 63.2"; // Speed 2 / Speed 0.0
//;
      A     #BRAKE_RELEASE_OK; // Release Brake - Confirm
      JCN   END;
      =     "A 63.1"; // Speed 1
      R     "A 63.2"; // Speed 2 = Off
      =     "A 63.3"; // H = Reverse (Dn)
      JU    END;
NETWORK
TITLE =Drive Off
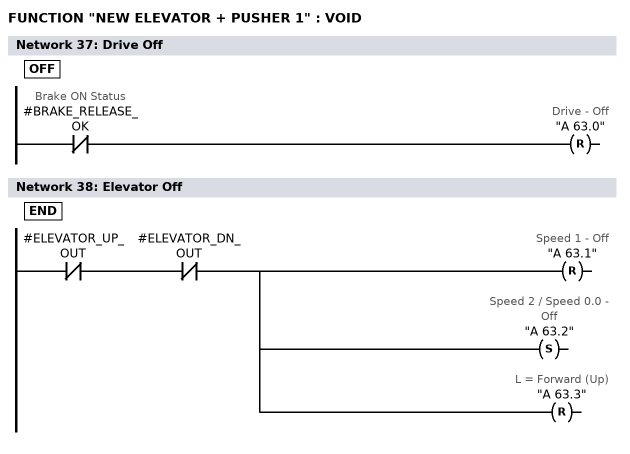

OFF:  AN    #BRAKE_RELEASE_OK; // Brake ON Status
      R     "A 63.0"; // Drive - Off
NETWORK
TITLE =Elevator Off

END:  AN    #ELEVATOR_UP_OUT;
      AN    #ELEVATOR_DN_OUT;
      R     "A 63.1"; // Speed 1 - Off
      S     "A 63.2"; // Speed 2 / Speed 0.0 - Off
      R     "A 63.3"; // L = Forward (Up)
END_FUNCTION

FUNCTION "NEW C1 - BELT" : VOID
TITLE =NEW FC918 (was FC1018) - Conveyor 1 Pos. 1
//
NAME : POS_3
VERSION : 0.0


VAR_TEMP
  MAIN_SERVICE_1_SW : BOOL ;
  SERVICE_RUN : BOOL ;
  INITIALISATION : BOOL ;
  SENSOR_TEST : BOOL ;
END_VAR
BEGIN
NETWORK
TITLE =Service Test

      A     "HMI_DB".ALL_SERVICE_ENABLE_SW;
      A     "HMI_DB".CONVEYOR_1_SERVICE_SW;
      A     "HMI_DB".SERVICE_SW_1_STATUS;
      =     #MAIN_SERVICE_1_SW;
//;
      A     #MAIN_SERVICE_1_SW;
      O     "M 18.1";
      JNB   CON1;
      A     "HMI_DB".HMI_CONVEYOR_1_TEST_SSW;
      =     #SERVICE_RUN;
      S     "DB UTILITY".Elevator_Disable;
      S     "DB UTILITY".Pusher_1_Disable;
//;
      A     "HMI_DB".SERVICE_INIT_PB;
      =     #INITIALISATION;
//;
      AN    #MAIN_SERVICE_1_SW;
      R     "HMI_DB".HMI_CONVEYOR_1_TEST_SSW;
      R     "DB UTILITY".Elevator_Disable;
      R     "DB UTILITY".Pusher_1_Disable;

CON1: R     #SERVICE_RUN;
      R     #INITIALISATION;
      FP    "FP 158.2";
      =     "M 18.1";
NETWORK
TITLE =Step 2N1 - Power ON
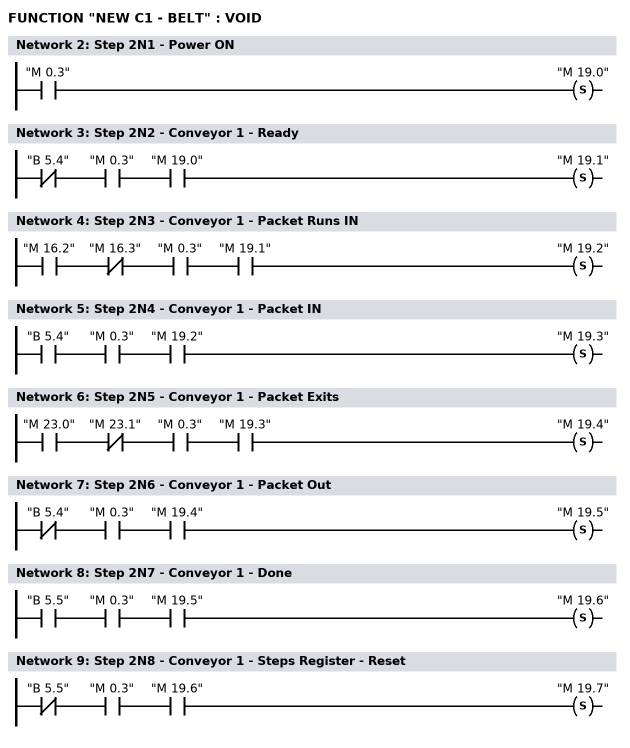

      A     "M 0.3";
      S     "M 19.0";
NETWORK
TITLE =Step 2N2 - Conveyor 1 - Ready

      AN    "B 5.4";
      A     "M 0.3";
      A     "M 19.0";
      S     "M 19.1";
NETWORK
TITLE =Step 2N3 - Conveyor 1 - Packet Runs IN

      A     "M 16.2";
      AN    "M 16.3";
      A     "M 0.3";
      A     "M 19.1";
      S     "M 19.2";
NETWORK
TITLE =Step 2N4 - Conveyor 1 - Packet IN

      A     "B 5.4";
      A     "M 0.3";
      A     "M 19.2";
      S     "M 19.3";
NETWORK
TITLE =Step 2N5 - Conveyor 1 - Packet Exits

      A     "M 23.0";
      AN    "M 23.1";
      A     "M 0.3";
      A     "M 19.3";
      S     "M 19.4";
NETWORK
TITLE =Step 2N6 - Conveyor 1 - Packet Out

      AN    "B 5.4";
      A     "M 0.3";
      A     "M 19.4";
      S     "M 19.5";
NETWORK
TITLE =Step 2N7 - Conveyor 1 - Done

      A     "B 5.5";
      A     "M 0.3";
      A     "M 19.5";
      S     "M 19.6";
NETWORK
TITLE =Step 2N8 - Conveyor 1 - Steps Register - Reset

      AN    "B 5.5";
      A     "M 0.3";
      A     "M 19.6";
      S     "M 19.7";
NETWORK
TITLE =Conveyor 1 - Steps Register - Reset

      A(    ;
      O     "M 19.7";
      O     "DB UTILITY".T19_DN;
      O     #INITIALISATION;
      O     "DB UTILITY".Conveyor_1_Disable;
      )     ;
      A     "M 0.3";
      JNB   INIT;
      L     W#16#0;
      T     "MW 19";

INIT: CLR   ;
NETWORK
TITLE =Soft Timer 19 Reset

      A     "M 19.2";
      AN    "M 19.3";
      A     "M 0.3";
      JCN   R191;
      JU    E191;

R191: L     L#0;
      T     "DB UTILITY".T19_ET;
      R     "DB UTILITY".T19_DN;

E191: NOP   0;

NETWORK
TITLE =Soft Timer 19 Add

      A     "M 19.2";
      AN    "M 19.3";
      A     "M 0.3";
      AN    "DB UTILITY".Freeze_Sequence_1;
      AN    "DB UTILITY".T19_DN;
      JCN   E192;

      L     "DB UTILITY".T19_ET;
      L     "DB UTILITY".Scan_Cycle_Previous;
      ITD   ;
      +D    ;
      T     "DB UTILITY".T19_ET;

E192: NOP   0;

NETWORK
TITLE =Soft Timer 19 Done 10s
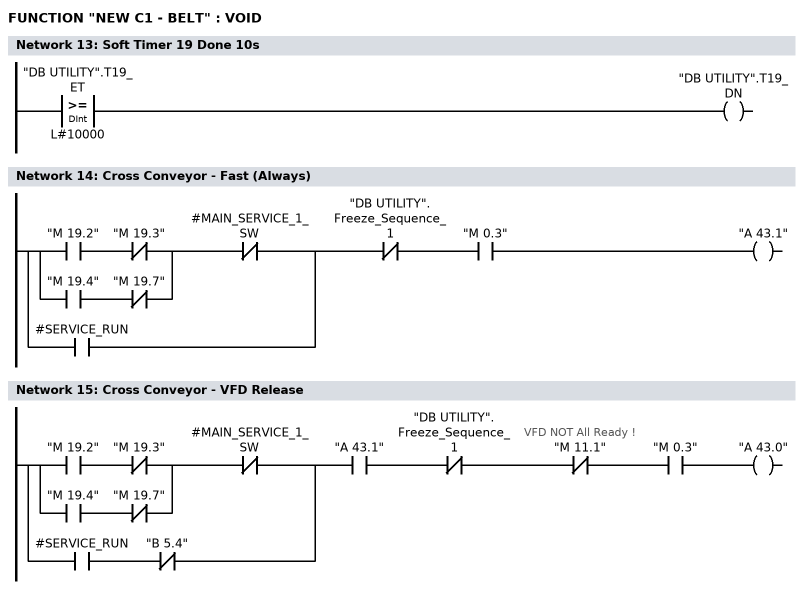

      L     "DB UTILITY".T19_ET;
      L     L#10000;
      >=D   ;
      =     "DB UTILITY".T19_DN;
NETWORK
TITLE =Cross Conveyor - Fast (Always)

      A(    ;
      A     "M 19.2";
      AN    "M 19.3";
      O     ;
      A     "M 19.4";
      AN    "M 19.7";
      )     ;
      AN    #MAIN_SERVICE_1_SW;
      O     #SERVICE_RUN;
      AN    "DB UTILITY".Freeze_Sequence_1;
      A     "M 0.3";
      =     "A 43.1";

NETWORK
TITLE =Cross Conveyor - VFD Release

      A(    ;
      A     "M 19.2";
      AN    "M 19.3";
      O     ;
      A     "M 19.4";
      AN    "M 19.7";
      )     ;
      AN    #MAIN_SERVICE_1_SW;
      O(    ;
      A     #SERVICE_RUN;
      AN    "B 5.4";
      )     ;
      A     "A 43.1";
      AN    "DB UTILITY".Freeze_Sequence_1;
      AN    "M 11.1"; // VFD NOT All Ready !
      A     "M 0.3";
      =     "A 43.0";
NETWORK
TITLE =Any Conveyors Packet mS Test
//    A     "B 10.7"
//    A     "A 48.6"
      A     "B 10.6";
      A     "A 48.3";






      =     #SENSOR_TEST;
//;
      A     #SENSOR_TEST;
      FP    "FP 147.7";
      JNB   NRST;
      L     0;
      T     "COLLATORS DB".Any_Conveyors_mS;

NRST: A     #SENSOR_TEST;
      JNB   NCNT;
      L     "COLLATORS DB".Any_Conveyors_mS;
      L     "DB UTILITY".Scan_Cycle_Previous;
      ITD   ;
      +D    ;
      T     "COLLATORS DB".Any_Conveyors_mS;

NCNT: CLR   ;

END_FUNCTION

FUNCTION "NEW C2 - ANGLE B+R" : VOID
TITLE =NEW FC922 (was FC1022) - Angle Conveyor 2 Pos. 4
NAME : POS_4
VERSION : 0.0


VAR_TEMP
  MAIN_SERVICE_1_SW : BOOL ;
  SERVICE_BELT_RUN : BOOL ;
  SERVICE_ROLLER_LIFT : BOOL ;
  SERVICE_ROLLER_RUN : BOOL ;
  INITIALISATION : BOOL ;
  PACKET_MEASURE_FLAG : BOOL ;
END_VAR
BEGIN
NETWORK
TITLE =Service Test

      A     "HMI_DB".ALL_SERVICE_ENABLE_SW;
      A     "HMI_DB".CONVEYOR_2_SERVICE_SW;
      A     "HMI_DB".SERVICE_SW_1_STATUS;
      =     #MAIN_SERVICE_1_SW;
//;
      A     #MAIN_SERVICE_1_SW;
      O     "M 22.1";
      JNB   CON2;
      A     "HMI_DB".HMI_CONVEYOR_2B_TEST_SSW;
      =     #SERVICE_BELT_RUN;
      S     "DB UTILITY".Conveyor_1_Disable;
//;
      A     "HMI_DB".HMI_CONVEYOR_2L_TEST_SSW;
      =     #SERVICE_ROLLER_LIFT;
      S     "DB UTILITY".Conveyor_1_Disable;
//;
      A     "HMI_DB".HMI_CONVEYOR_2R_TEST_SSW;
      =     #SERVICE_ROLLER_RUN;
      S     "DB UTILITY".Conveyor_1_Disable;
//;
      A     "HMI_DB".SERVICE_INIT_PB;
      =     #INITIALISATION;
//;
      AN    #MAIN_SERVICE_1_SW;
      R     "HMI_DB".HMI_CONVEYOR_2B_TEST_SSW;
      R     "HMI_DB".HMI_CONVEYOR_2L_TEST_SSW;
      R     "HMI_DB".HMI_CONVEYOR_2R_TEST_SSW;
      R     "DB UTILITY".Conveyor_1_Disable;

CON2: R     #SERVICE_BELT_RUN;
      R     #SERVICE_ROLLER_LIFT;
      R     #SERVICE_ROLLER_RUN;
      R     #INITIALISATION;
      FP    "FP 158.3";
      =     "M 22.1";

NETWORK
TITLE =Angle Conveyor - Fault / Ready
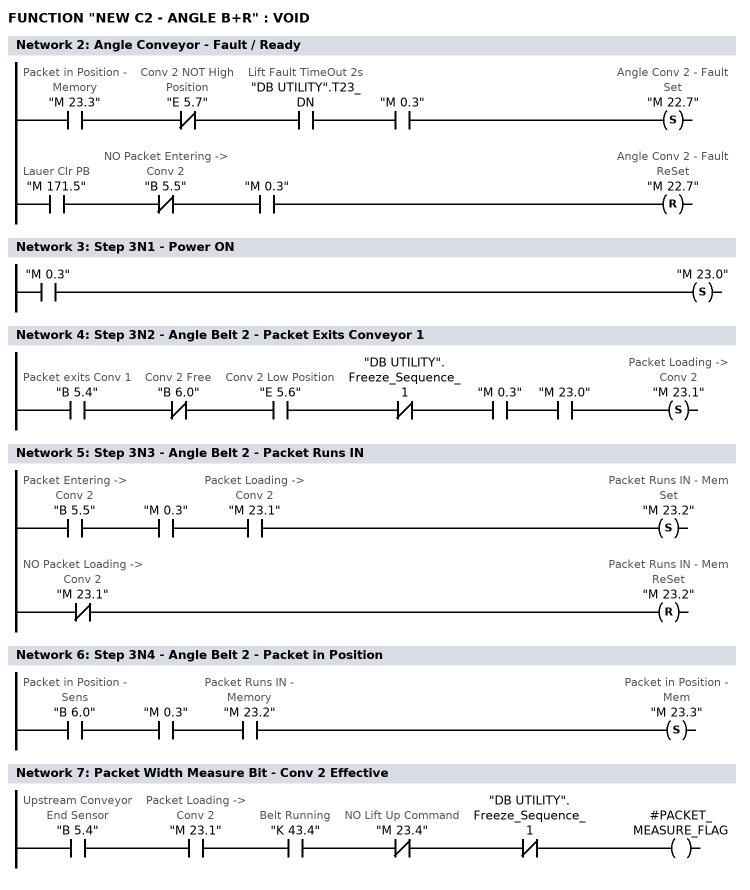

      A     "M 23.3"; // Packet in Position - Memory
      AN    "E 5.7"; // Conv 2 NOT High Position
      A     "DB UTILITY".T23_DN; // Lift Fault TimeOut 2s
      A     "M 0.3";
      S     "M 22.7"; // Angle Conv 2 - Fault Set
//;
      A     "M 171.5"; // Lauer Clr PB
      AN    "B 5.5"; // NO Packet Entering -> Conv 2
      A     "M 0.3";
      R     "M 22.7"; // Angle Conv 2 - Fault ReSet

NETWORK
TITLE =Step 3N1 - Power ON

      A     "M 0.3";
      S     "M 23.0";

NETWORK
TITLE =Step 3N2 - Angle Belt 2 - Packet Exits Conveyor 1

      A     "B 5.4"; // Packet exits Conv 1
      AN    "B 6.0"; // Conv 2 Free
      A     "E 5.6"; // Conv 2 Low Position
      AN    "DB UTILITY".Freeze_Sequence_1;
      A     "M 0.3";
      A     "M 23.0";
      S     "M 23.1"; // Packet Loading -> Conv 2
NETWORK
TITLE =Step 3N3 - Angle Belt 2 - Packet Runs IN

      A     "B 5.5"; // Packet Entering -> Conv 2
      A     "M 0.3";
      A     "M 23.1"; // Packet Loading -> Conv 2
      S     "M 23.2"; // Packet Runs IN - Mem Set
//;
      ON    "M 23.1"; // NO Packet Loading -> Conv 2
      R     "M 23.2"; // Packet Runs IN - Mem ReSet

NETWORK
TITLE =Step 3N4 - Angle Belt 2 - Packet in Position

      A     "B 6.0"; // Packet in Position - Sens
      A     "M 0.3";
      A     "M 23.2"; // Packet Runs IN - Memory
      S     "M 23.3"; // Packet in Position - Mem
NETWORK
TITLE =Packet Width Measure Bit - Conv 2 Effective

      A     "B 5.4"; // Upstream Conveyor End Sensor
      A     "M 23.1"; // Packet Loading -> Conv 2
      A     "K 43.4"; // Belt Running
      AN    "M 23.4"; // NO Lift Up Command
      AN    "DB UTILITY".Freeze_Sequence_1;
      =     #PACKET_MEASURE_FLAG;

NETWORK
TITLE =Packet Width Time Reset - Freeze Safe

      A     "M 23.1"; // Packet Loading -> Conv 2
      O     "DB UTILITY".Freeze_Sequence_1;
      JC    NRS1;

      L     L#0;
      T     "MD 260"; // Width [mS]

NRS1: NOP   0;
NETWORK
TITLE =Packet Width Time Count Up From Sensor "B 5.4"

      A     #PACKET_MEASURE_FLAG;
      JCN   NMES;

      L     "MD 260"; // Width [mS]
      L     "DB UTILITY".Scan_Cycle_Previous;
      ITD   ;
      +D    ;
      T     "MD 260"; // Width [mS]

NMES: NOP   0;
NETWORK
TITLE =Middle Travel Time Reset - Freeze Safe

      A     "M 23.3"; // Packet in Position - Mem
      O     "DB UTILITY".Freeze_Sequence_1;
      JC    NRS2;

      L     L#0;
      T     "MD 264"; // Half Width [mS] - Zeroed

NRS2: NOP   0;
NETWORK
TITLE =Middle Travel Time Count Up From B 6.0

      ON    "M 23.3"; // NO Packet in Position - Mem
      O     "M 23.4"; // Lift Up Command
      ON    "K 43.4"; // Belt Stopped
      ON    "M 0.3"; // No Power
      AN    "DB UTILITY".Freeze_Sequence_1;
      JC    NCNT;

      L     "MD 264"; // Half Width [mS]
      L     "DB UTILITY".Scan_Cycle_Previous;
      ITD   ;
      +D    ;
      T     "MD 264"; // Half Width [mS] - Add

NCNT: NOP   0;
NETWORK
TITLE =Middle Travel Time Clamp Zero

      L     "MD 264"; // Half Width [mS]
      L     L#0;
      >=D   ;
      JC    NMID;

      L     L#0;
      T     "MD 264"; // Half Width [mS] - Reset

NMID: NOP   0;
NETWORK
TITLE =Soft Timer 23 Reset - Lift Fault TimeOut 2s + Freeze Option

      A     "M 23.3"; // Packet in Position - Memory
      AN    "M 23.4"; // NO Lift Up Command
      A     "M 0.3";
      JCN   R231;
      JU    E231;

R231: L     L#0;
      T     "DB UTILITY".T23_ET;
      R     "DB UTILITY".T23_DN;

E231: NOP   0;

NETWORK
TITLE =Soft Timer 23 Add

      A     "M 23.3"; // Packet in Position - Memory
      AN    "M 23.4"; // NO Lift Up Command
      A     "M 0.3";
      AN    "DB UTILITY".Freeze_Sequence_1; // Sequence Freezer Bit
      AN    "DB UTILITY".T23_DN;
      JCN   E232;

      L     "DB UTILITY".T23_ET;
      L     "DB UTILITY".Scan_Cycle_Previous;
      ITD   ;
      +D    ;
      T     "DB UTILITY".T23_ET;

E232: NOP   0;

NETWORK
TITLE =Soft Timer 23 Done 2s

      L     "DB UTILITY".T23_ET;
      L     L#2500; // [mS]
      >=D   ;
      =     "DB UTILITY".T23_DN;
NETWORK
TITLE =Soft Timer 24 Reset - Belt TimeOut 8s + Freeze Option

      A     "M 23.1";
      AN    "M 23.3";
      A     "K 43.4";
      A     "M 0.3";
      JCN   R241;
      JU    E241;

R241: L     L#0;
      T     "DB UTILITY".T24_ET;
      R     "DB UTILITY".T24_DN;

E241: NOP   0;

NETWORK
TITLE =Soft Timer 24 Add

      A     "M 23.1";
      AN    "M 23.3";
      A     "K 43.4";
      A     "M 0.3";
      AN    "DB UTILITY".Freeze_Sequence_1;
      AN    "DB UTILITY".T24_DN;
      JCN   E242;

      L     "DB UTILITY".T24_ET;
      L     "DB UTILITY".Scan_Cycle_Previous;
      ITD   ;
      +D    ;
      T     "DB UTILITY".T24_ET;

E242: NOP   0;

NETWORK
TITLE =Soft Timer 24 Done 8s

      L     "DB UTILITY".T24_ET;
      L     L#8000;
      >=D   ;
      =     "DB UTILITY".T24_DN;
      S     "M 24.4";
NETWORK
TITLE =Step 3N5 - Angle Belt - Lift ("MD 264" to Center the Packet)

      A(    ;
      A(    ;
      L     "MD 264";
      L     L#2;
      *D    ;
      L     "MD 260";
      >=D   ;
      )     ;
      AN    #PACKET_MEASURE_FLAG;
      AN    "B 5.5";
      O     "DB UTILITY".T23_DN;
      )     ;
      A     "M 0.3";
      A     "M 23.3";
      S     "M 23.4";
NETWORK
TITLE =Step 3N6 - Angle Rollers - Up
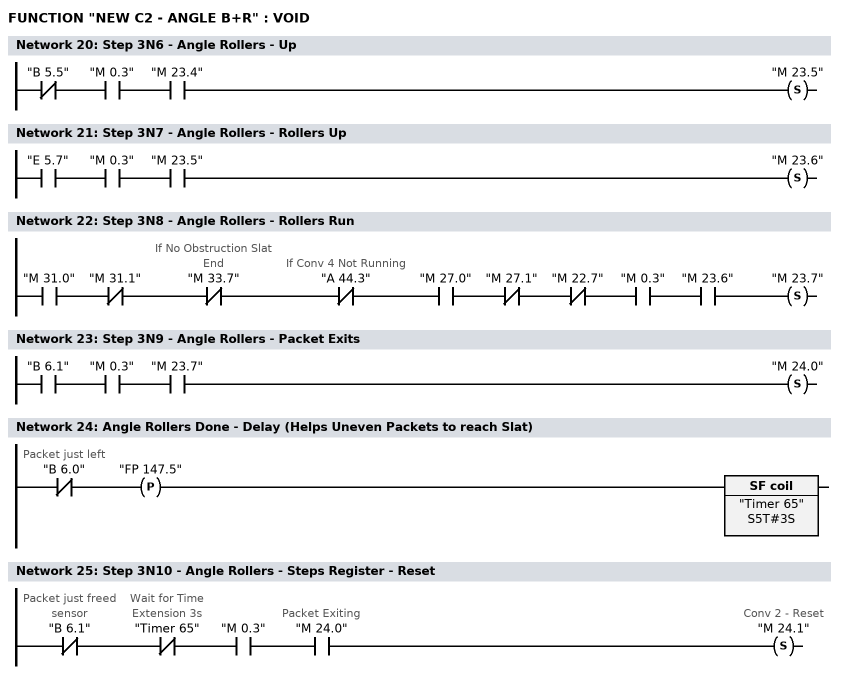

      AN    "B 5.5";
      A     "M 0.3";
      A     "M 23.4";
      S     "M 23.5";

NETWORK
TITLE =Step 3N7 - Angle Rollers - Rollers Up

      A     "E 5.7";
      A     "M 0.3";
      A     "M 23.5";
      S     "M 23.6";

NETWORK
TITLE =Step 3N8 - Angle Rollers - Rollers Run

      A     "M 31.0";
      AN    "M 31.1";
      AN    "M 33.7"; // If No Obstruction Slat End
      AN    "A 44.3"; // If Conv 4 Not Running
      A     "M 27.0";
      AN    "M 27.1";
      AN    "M 22.7";
      A     "M 0.3";
      A     "M 23.6";
      S     "M 23.7";

NETWORK
TITLE =Step 3N9 - Angle Rollers - Packet Exits

      A     "B 6.1";
      A     "M 0.3";
      A     "M 23.7";
      S     "M 24.0";

NETWORK
TITLE =Angle Rollers Done - Delay (Helps Uneven Packets to reach Slat)

      AN    "B 6.0"; // Packet just left
      FP    "FP 147.5";
      L     S5T#3S;
      SF    "Timer 65"; // Time Extension 3s
NETWORK
TITLE =Step 3N10 - Angle Rollers - Steps Register - Reset

      AN    "B 6.1"; // Packet just freed sensor
      AN    "Timer 65"; // Wait for Time Extension 3s
      A     "M 0.3";
      A     "M 24.0"; // Packet Exiting
      S     "M 24.1"; // Conv 2 - Reset
NETWORK
TITLE =Conveyor 2 - Steps Register - Reset

      A(    ;
      O     "M 24.1";
      O     "DB UTILITY".T24_DN;
      O     "DB UTILITY".T25_DN;
      O     #INITIALISATION;
      O     "DB UTILITY".Conveyor_1_Disable;
      )     ;
      A     "M 0.3";
      JC    M001;
      JU    M002;

M001: L     W#16#0;
      T     "MW 23";

M002: NOP   0;
NETWORK
TITLE =Soft Timer 25 Reset - Roller TimeOut 8s + Freeze Option

      A     "M 23.7";
      AN    "M 24.1";
      A     "M 0.3";
      JCN   R251;
      JU    E251;

R251: L     L#0;
      T     "DB UTILITY".T25_ET;
      R     "DB UTILITY".T25_DN;

E251: NOP   0;

NETWORK
TITLE =Soft Timer 25 Add

      A     "M 23.7";
      AN    "M 24.1";
      A     "M 0.3";
      AN    "DB UTILITY".Freeze_Sequence_2;
      AN    "DB UTILITY".T25_DN;
      JCN   E252;

      L     "DB UTILITY".T25_ET;
      L     "DB UTILITY".Scan_Cycle_Previous;
      ITD   ;
      +D    ;
      T     "DB UTILITY".T25_ET;

E252: NOP   0;

NETWORK
TITLE =Soft Timer 25 Done 8s

      L     "DB UTILITY".T25_ET;
      L     L#8000;
      >=D   ;
      =     "DB UTILITY".T25_DN;
NETWORK
TITLE =Angle Conveyor Belt - Run

      A     "M 23.1";
      AN    "M 23.4";
      AN    #MAIN_SERVICE_1_SW;
      O(    ;
      A     #SERVICE_BELT_RUN;
      A(    ;
      A     "B 6.0";
      L     S5T#200MS;
      SD    "Timer 21";
//;
      AN    "Timer 21";
      )     ;
      )     ;
      AN    "M 22.7";
      AN    "DB UTILITY".Freeze_Sequence_1;
      AN    "M 11.1"; // VFD NOT All Ready !
      A     "M 0.3";
      =     "K 43.4";

NETWORK
TITLE =Angle Conveyor Rollers - Run
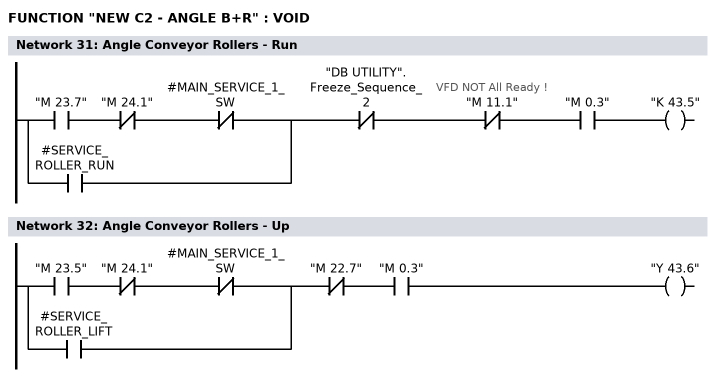

      A     "M 23.7";
      AN    "M 24.1";
      AN    #MAIN_SERVICE_1_SW;
      O     #SERVICE_ROLLER_RUN;
      AN    "DB UTILITY".Freeze_Sequence_2;
      AN    "M 11.1"; // VFD NOT All Ready !
      A     "M 0.3";
      =     "K 43.5";

NETWORK
TITLE =Angle Conveyor Rollers - Up

      A     "M 23.5";
      AN    "M 24.1";
      AN    #MAIN_SERVICE_1_SW;
      O     #SERVICE_ROLLER_LIFT;
      AN    "M 22.7";
      A     "M 0.3";
      =     "Y 43.6";
END_FUNCTION

FUNCTION "NEW C3 - SLAT PIW" : VOID
TITLE =FC 925 > NEW FC924 (was FC1024) - Slat Conveyor 3 Pos.5
//v0.1 2026-11-19: C3 encoder Ch0 read DIRECT every scan: PIW 328 (HW Config
//User_Type1 right) instead of "FM350 DB".ACT_CNTV0 (read job, ~100 mS old).
NAME : POS_5
VERSION : 0.1


VAR_TEMP
  MAIN_SERVICE_1_SW : BOOL ;
  SERVICE_RUN : BOOL ;
  INITIALISATION : BOOL ;
END_VAR
BEGIN
NETWORK
TITLE =Service Test

      A     "HMI_DB".ALL_SERVICE_ENABLE_SW;
      A     "HMI_DB".CONVEYOR_3_SERVICE_SW;
      A     "HMI_DB".SERVICE_SW_1_STATUS;
      =     #MAIN_SERVICE_1_SW;
//;
      A     #MAIN_SERVICE_1_SW;
      O     "M 26.3";
      JNB   CON3;
      A     "HMI_DB".HMI_CONVEYOR_3_TEST_SSW;
      =     #SERVICE_RUN;
      S     "DB UTILITY".Conveyor_2_Disable;
//;
      AN    #MAIN_SERVICE_1_SW;
      R     "HMI_DB".HMI_CONVEYOR_3_TEST_SSW;
      R     "DB UTILITY".Conveyor_2_Disable;
//;
      A     "HMI_DB".SERVICE_INIT_PB;
      A     #MAIN_SERVICE_1_SW;
      =     #INITIALISATION;

CON3: R     #SERVICE_RUN;
      R     #INITIALISATION; // Fix: temp not written when service is off
      FP    "FP 227.0";
      =     "M 26.3";
NETWORK
TITLE =Packet Length Measurements [mm] - While Collating

      A     "B 6.2"; // C3 InFeed Sens - New Packet
      FP    "FP 227.1";
      A     "A 44.0";
      JC    PRNT;
      JU    RPRT;

PRNT: L     "PIW 328"; // Direct Ch0 (was ACT_CNTV0, ~100 mS old)
      T     "HOUSE_KEEPING DB".C3_Encoder_READ_Mem;

RPRT: AN    "B 6.2"; // C3 InFeed Sens - New Packet End
      FP    "FP 227.2";
      JCN   NTKE;

      L     "PIW 328"; // Direct Ch0 (was ACT_CNTV0, ~100 mS old)
      L     "HOUSE_KEEPING DB".C3_Encoder_READ_Mem;
      -I    ;
      T     "HOUSE_KEEPING DB".C3_Packet_Length_ep;
      DTR   ;
//;
      L     1.300000e+000; //  Encoder Wheel 900mm / 600 PPR  [mm/pulse]
      *R    ;
      RND   ;
      T     "HOUSE_KEEPING DB".C3_Packet_Length_mm;

NTKE: NOP   0;
NETWORK
TITLE =Slat Conveyor 3 - Packets / Conveyor Length - Calculation

      A     "M 27.1";
      FP    "FP 227.3";
      JNB   M271;
      L     "COLLATORS DB".Conveyor_Length_C3;
      ITD   ;
      DTR   ;
      L     5.000000e+000;
      /R    ;
      RND   ;
      T     "COLLATORS DB".Press_Length_C3;
      T     "MW 212";

M271: NOP   0;
NETWORK
TITLE =Slat Conveyor 3 - Surface Length Manager (PulseUnit)

      A     "M 27.1";
      O     "M 26.6";
      S     "M 166.0";
//;
      A     "M 166.0";
      O(    ;
      AN    "M 10.0";
      FP    "FP 227.4";
      )     ;
      =     "FM350 DB".CONTROL_SIGNALS.SW_GATE0; // C3 Surface Count
//;
      A     "M 166.0"; // Start Count (100mS Pulse)
      A(    ;
      L     "PIW 328"; // Direct Ch0 (was ACT_CNTV0, ~100 mS old) C3 Surface Count
      L     "MW 212";
      >=I   ;
      )     ;
      A     "M 0.3";
      JCN   R291;
      JU    E291;

R291: L     L#0;
      T     "DB UTILITY".T27_ET;
      R     "DB UTILITY".T27_DN;

E291: NOP   0;
NETWORK
TITLE =Soft Timer 27 Add - FM350 needs a 100mS Pulse !

      A     "M 166.0";
      A(    ;
      L     "PIW 328"; // Direct Ch0 (was ACT_CNTV0, ~100 mS old) C3 Surface Count
      L     "MW 212";
      >=I   ;
      )     ;
      A     "M 0.3";
      AN    "DB UTILITY".Freeze_Sequence_2;
      AN    "DB UTILITY".T27_DN;
      JCN   E292;

      L     "DB UTILITY".T27_ET;
      L     "DB UTILITY".Scan_Cycle_Previous;
      ITD   ;
      +D    ;
      T     "DB UTILITY".T27_ET;

E292: NOP   0;
NETWORK
TITLE =Soft Timer 27 Done 100mS  // Start Count (100mS Pulse)
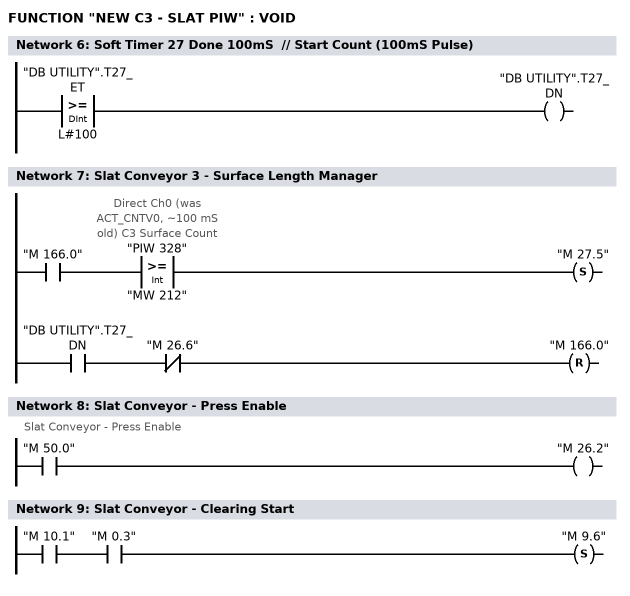

      L     "DB UTILITY".T27_ET;
      L     L#100;
      >=D   ;
      =     "DB UTILITY".T27_DN;
NETWORK
TITLE =Slat Conveyor 3 - Surface Length Manager

      A     "M 166.0";
      A(    ;
      L     "PIW 328"; // Direct Ch0 (was ACT_CNTV0, ~100 mS old) C3 Surface Count
      L     "MW 212";
      >=I   ;
      )     ;
      S     "M 27.5";
//;
      A     "DB UTILITY".T27_DN;
      AN    "M 26.6";
      R     "M 166.0";
NETWORK
TITLE =Slat Conveyor - Press Enable
//Slat Conveyor - Press Enable
      A     "M 50.0";
      =     "M 26.2";
NETWORK
TITLE =Slat Conveyor - Clearing Start

      A     "M 10.1";
      A     "M 0.3";
      S     "M 9.6";
NETWORK
TITLE =Slat Conveyor - Clearing
//Counting 9K Pulses Should Suffice !
      A     "M 10.1";
      AN    "M 10.2";
      AN    "A 44.0";
      S     "M 26.6";
//;
      A     "M 26.6";
      JNB   M266;
      A(    ;
      L     "PIW 328"; // Direct Ch0 (was ACT_CNTV0, ~100 mS old) C3 Surface Count
      L     10000;
      >I    ;
      )     ;
      =     "M 26.7";

M266: NOP   0;

      A     "M 26.7";
      ON    "M 10.0";
      R     "M 26.6";
NETWORK
TITLE =Slat Conveyor Steps
//Slat Conveyor Steps


NETWORK
TITLE =Step 4N1 - Power ON
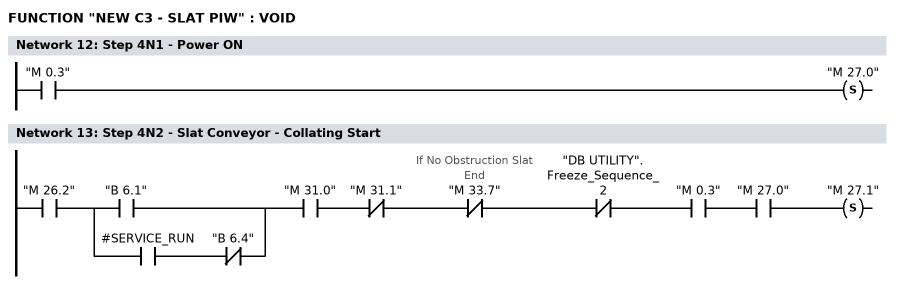

      A     "M 0.3";
      S     "M 27.0";
NETWORK
TITLE =Step 4N2 - Slat Conveyor - Collating Start

      A     "M 26.2";
      A(    ;
      O     "B 6.1";
      O(    ;
      A     #SERVICE_RUN;
      AN    "B 6.4";
      )     ;
      )     ;
      A     "M 31.0";
      AN    "M 31.1";
      AN    "M 33.7"; // If No Obstruction Slat End
      AN    "DB UTILITY".Freeze_Sequence_2;
      A     "M 0.3";
      A     "M 27.0";
      S     "M 27.1";
NETWORK
TITLE =Soft Timer 28 Reset - Collating TimeOut + Freeze Option

      A     "M 27.1";
      AN    "M 27.4";
      A     "M 0.3";
      JCN   R271;
      JU    E271;

R271: L     L#0;
      T     "DB UTILITY".T28_ET;
      R     "DB UTILITY".T28_DN;

E271: NOP   0;
NETWORK
TITLE =Soft Timer 28 Add

      A     "M 27.1";
      AN    "M 27.4";
      A     "M 0.3";
      AN    "DB UTILITY".Freeze_Sequence_2;
      AN    "DB UTILITY".T28_DN;
      JCN   E272;

      L     "DB UTILITY".T28_ET;
      L     "DB UTILITY".Scan_Cycle_Previous;
      ITD   ;
      +D    ;
      T     "DB UTILITY".T28_ET;

E272: NOP   0;
NETWORK
TITLE =Soft Timer 27 Done 11s
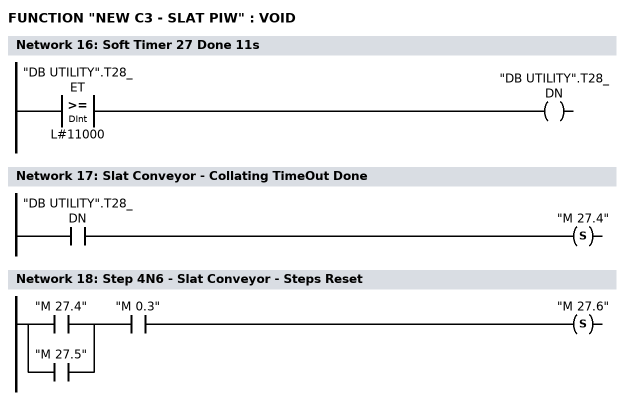

      L     "DB UTILITY".T28_ET;
      L     L#11000;
      >=D   ;
      =     "DB UTILITY".T28_DN;
NETWORK
TITLE =Slat Conveyor - Collating TimeOut Done

      A     "DB UTILITY".T28_DN;
      S     "M 27.4";
NETWORK
TITLE =Step 4N6 - Slat Conveyor - Steps Reset

      O     "M 27.4";
      O     "M 27.5";
      A     "M 0.3";
      S     "M 27.6";
NETWORK
TITLE =Slat Conveyor - Steps Register - Reset

      A(    ;
      O     "M 27.6";
      O     #INITIALISATION;
      O     "DB UTILITY".Conveyor_3_Disable;
      )     ;
      A     "M 0.3";
      JC    M001;
      JU    M002;

M001: L     W#16#0;
      T     "MB 27";
      R     "M 26.7";

M002: NOP   0;
NETWORK
TITLE =Slat Conveyor - VFD Release

      A(    ;
      O     "M 27.1";
      O     "M 26.6";
      )     ;
      AN(   ;
      A     "M 26.6";
      A     "M 31.5";
      )     ;
      AN    "DB UTILITY".Freeze_Sequence_2;
      AN    "M 11.1"; // VFD NOT All Ready !
      A     "M 0.3";
      =     "A 44.0";
      =     "A 44.1";
END_FUNCTION

FUNCTION "NEW C4 - COLLATOR PIW" : VOID
TITLE =FC 932 > NEW FC931 (was FC1031) - Collator Conveyor 4 Pos.6
//Collator Conveyor 4 - Is On Both Service Pages 1 & 2
//v0.1 2026-11-19: C4 encoders read DIRECT every scan: Ch2 = PIW 332, Ch3 = PIW
//330
//(HW Config) instead of ACT_CNTV2/3 (read job, ~100 mS old).
NAME : POS_6
VERSION : 0.1


VAR_TEMP
  MAIN_SERVICE_1_2_SW : BOOL ;	//Collator Conveyor 4 - On Service 1 & 2
  SERVICE_RUN : BOOL ;
  INITIALISATION : BOOL ;
  COUNTER_TRIGGER : BOOL ;
  PACKET_LENGTH_4 : WORD ;	//Collator Conveyor 4 - Packet Length
  W_TUBE_mm : WORD ;
  W_TUBE_PERCENT : WORD ;	//Tube 5 % Value
  R_TUBE_PERCENT : REAL ;	//Tube 5 % Value
  R_TUBE_mm : REAL ;
END_VAR
BEGIN
NETWORK
TITLE =Conveyor 4 - Service

      A     "HMI_DB".ALL_SERVICE_ENABLE_SW;
      A     "HMI_DB".CONVEYOR_4_SERVICE_SW;
      A(    ;
      O     "HMI_DB".SERVICE_SW_1_STATUS;
      O     "HMI_DB".SERVICE_SW_2_STATUS;
      )     ;
      =     "HMI_DB".SERVICE_SW_1_2_STATUS;
      =     #MAIN_SERVICE_1_2_SW;
//;
      A     #MAIN_SERVICE_1_2_SW;
      O     "M 26.1";
      JNB   CON4;
      A     "HMI_DB".HMI_CONVEYOR_4_TEST_SSW;
      =     #SERVICE_RUN;
      S     "DB UTILITY".Conveyor_3_Disable;
//;
      A     "HMI_DB".SERVICE_INIT_PB;
      A     #MAIN_SERVICE_1_2_SW;
      =     #INITIALISATION;
//;
      AN    #MAIN_SERVICE_1_2_SW;
      R     "HMI_DB".HMI_CONVEYOR_4_TEST_SSW;
      R     "DB UTILITY".Conveyor_3_Disable;

CON4: R     #SERVICE_RUN;
      R     #INITIALISATION;
      FP    "FP 158.4";
      =     "M 26.1";
NETWORK
TITLE =Soft Timer 90 Reset Conveyor 4 - Encoder has Stop L - Timer  500

      AN    "E 6.6";
      AN    "M 30.0";
      A     "M 0.3";
      JCN   R900;
      JU    E900;

R900: L     L#0;
      T     "DB UTILITY".T90_ET;
      R     "DB UTILITY".T90_DN;

E900: NOP   0;
NETWORK
TITLE =Soft Timer 90 Add Conveyor 4 - Encoder has Stop H - Timer  500mS

      AN    "E 6.6";
      AN    "M 30.0";
      A     "M 0.3";
      AN    "DB UTILITY".Freeze_Sequence_2;
      AN    "DB UTILITY".T90_DN;
      JCN   E901;

      L     "DB UTILITY".T90_ET;
      L     "DB UTILITY".Scan_Cycle_Previous;
      ITD   ;
      +D    ;
      T     "DB UTILITY".T90_ET;

E901: NOP   0;
NETWORK
TITLE =Soft Timer 90 Done 500mS

      L     "DB UTILITY".T90_ET;
      L     L#500;
      >=D   ;
      =     "DB UTILITY".T90_DN;
NETWORK
TITLE =Soft Timer 91 Reset

      A     "E 6.6";
      AN    "M 30.0";
      A     "M 0.3";
      JCN   R910;
      JU    E910;

R910: L     L#0;
      T     "DB UTILITY".T91_ET;
      R     "DB UTILITY".T91_DN;

E910: NOP   0;
NETWORK
TITLE =Soft Timer 91 Add

      A     "E 6.6";
      AN    "M 30.0";
      A     "M 0.3";
      AN    "DB UTILITY".Freeze_Sequence_2;
      AN    "DB UTILITY".T91_DN;
      JCN   E911;

      L     "DB UTILITY".T91_ET;
      L     "DB UTILITY".Scan_Cycle_Previous;
      ITD   ;
      +D    ;
      T     "DB UTILITY".T91_ET;

E911: NOP   0;
NETWORK
TITLE =Soft Timer 91 Done 500mS
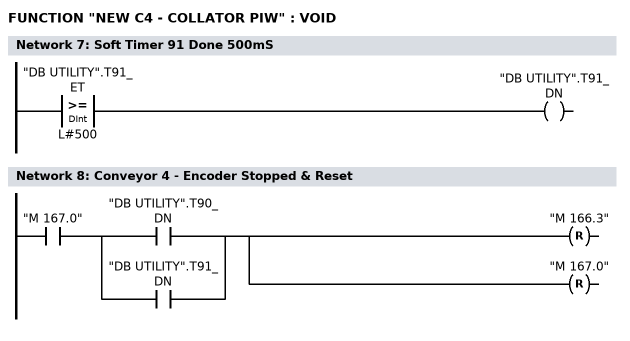

      L     "DB UTILITY".T91_ET;
      L     L#500;
      >=D   ;
      =     "DB UTILITY".T91_DN;
NETWORK
TITLE =Conveyor 4 - Encoder Stopped & Reset

      A     "M 167.0";
      A(    ;
      O     "DB UTILITY".T90_DN;
      O     "DB UTILITY".T91_DN;
      )     ;
      R     "M 166.3";
      R     "M 167.0";
NETWORK
TITLE =Conveyor 4 - Packet Length - Measurements

      A     "B 6.7";
      A     "M 31.1";
      S     "M 166.2"; // Counter 2 Gate - Set
      =     #COUNTER_TRIGGER;
//;
      A     "M 166.2"; // Counter 2
      =     "FM350 DB".CONTROL_SIGNALS.SW_GATE2; // C4 Length Count
//;
      A     "M 166.2"; // Counter 2
      O     "B 6.4";
      FP    "FP 149.4";
      JNB   NRAZ;
      L     0; // Reset First
      T     "COLLATORS DB".Packet_Length_C4_mS;

NRAZ: A     "M 166.2"; // Counter 2
      JNB   NCNT;
      L     "COLLATORS DB".Packet_Length_C4_mS;
      L     "DB UTILITY".Scan_Cycle_Previous;
      +I    ;
      T     "COLLATORS DB".Packet_Length_C4_mS; // Added ScanCycles

NCNT: A     "M 166.2"; // Counter 2
      AN    "B 6.4";
      AN    "B 6.7";
      JNB   B067;
      L     "PIW 332"; // Direct Ch2 (was ACT_CNTV2, ~100 mS old) C4 Length Count
      T     "COLLATORS DB".PacketLength_C4; // Encoder Pulses - Length
      T     #PACKET_LENGTH_4;
//;
      L     #PACKET_LENGTH_4;
      ITD   ;
      DTR   ;
      L     2.000000e-001;
      *R    ;
      RND   ;
      T     "COLLATORS DB".Frac_Packet_Length_C4;
//;
      L     #PACKET_LENGTH_4;
      +I    ;
      T     "COLLATORS DB".Packet_Length_Frac_C4;
      R     "M 166.2"; // Counter 2 Gate - Reset
      S     "M 167.1";
      S     "M 167.4";

B067: NOP   0;
NETWORK
TITLE =Packet Length Measurements [mm] - While Collating
//    A     "HOUSE_KEEPING DB".C4_First_Collating
      A     "B 6.7"; // C4 InFeed Sens - New Packet
      FP    "FP 226.1";
      A     "A 44.3";
      JCN   NPRT;

      L     "PIW 330"; // Direct Ch3 (was ACT_CNTV3, ~100 mS old)
      T     "HOUSE_KEEPING DB".C4_Encoder_READ_Mem;

NPRT: AN    "B 6.7"; // C4 InFeed Sens - New Packet End
      FP    "FP 226.2";
      JCN   NTKE;

      L     "PIW 330"; // Direct Ch3 (was ACT_CNTV3, ~100 mS old)
      L     "HOUSE_KEEPING DB".C4_Encoder_READ_Mem;
      -I    ;
      T     "HOUSE_KEEPING DB".C4_Packet_Length_ep; // C4 Packet Length [ep]
      DTR   ;
//;
      L     6.350000e+000; //  Encoder Wheel 635mm / 100 PPR  [mm/pulse]
      *R    ;
      RND   ;
      T     "HOUSE_KEEPING DB".C4_Packet_Length_mm;

NTKE: NOP   0;
NETWORK
TITLE =Packet Length Measurements [mS] - While Transfering to C5

      A     "M 31.6"; // C4 Transfer Step
      A     "B 7.0"; // C4 This Packet Exiting
      JCN   NMSR;
      L     "HOUSE_KEEPING DB".C4_Added_Scans_mS;
      L     "DB UTILITY".Scan_Cycle_Previous;
      +I    ;
      T     "HOUSE_KEEPING DB".C4_Added_Scans_mS; // Adding mS

NMSR: A     "M 31.6"; // C4 Transfer Step
      AN    "B 7.0"; // C4 This Packet Exiting Done
      FP    "FP 226.3";
      JCN   NLNT;

      L     "HOUSE_KEEPING DB".C4_Added_Scans_mS;
      T     "HOUSE_KEEPING DB".C4_Packet_Length_mS; // Packet Length mS @ 31 m/min
//;
      L     0;
      T     "HOUSE_KEEPING DB".C4_Added_Scans_mS; // Packet Length mS - Zeroed

NLNT: NOP   0;
NETWORK
TITLE =Between Packets Spaces - Measurements [mm]
